(* IEC 61131-3 sources: Masterarbeit/sigmatek/lasalclass2/PW022_hardware/Class/SafetyManager (part 5) *)

END_FUNCTION

FUNCTION MyXSort VAR_INPUT p1:^void; p2:^void; END_VAR VAR_OUTPUT retcode : dint; END_VAR;

FUNCTION SafetyManager::MySort
  VAR_INPUT
    src 	: ^USINT;
    no 	: UDINT;
    itemsize 	: UDINT;
    sortfunct 	: ^void;
  END_VAR
  VAR_OUTPUT
    retcode 	: BOOL;
  END_VAR
  var
    tmp, hp : ^DINT;
    mx, nx, wx, parent, child, max, i : dint;
    spuf : array[0..127] of dint;
  end_var

  retcode := false;

  // work faster with the pointer list (no memcopy used)
  if itemsize = 4 then
    nx      := to_dint(no);
    mx      := (nx + 6) / 8;
    src     := src;
    tmp     := #spuf[0];
    retcode := true;

    while(1) do
      if(mx) then
        mx     -= 1;
        parent := mx;
        tmp^ := (src$^DINT + (parent$udint*4))^;
      else
        nx -= 1;
        if(nx) then
          hp := src + (nx$udint*4);
          tmp^ := hp^;
          hp^ := (src$^DINT)^;
          parent := 0;
        else
          exit;
        end_if;
      end_if;

      child := parent * 8 + 1;
      while(child < nx) do
        wx := nx - child;
        if(wx > 8) then
          wx := 8;
        end_if;

        max := 0;
        if(wx > 1) then
          for i:=1 to wx-1 do
            if(sortfunct$MyXSort(src+(to_udint(child+i)*4), src+to_udint(child+max)*4) > 0) then
              max := i;
            end_if;
          end_for;
        end_if;

        child += max;

        if(sortfunct$MyXSort(src+(child$udint*4), tmp) <= 0) then
          exit;
        end_if;

        (src$^DINT+(parent$udint*4))^ := (src$^DINT+(child$udint*4))^;
        parent := child;
        child  := parent * 8 + 1;
      end_while;

      (src$^DINT+(parent$udint*4))^ := tmp^;
    end_while;
  else
    if(itemsize <= sizeof(spuf)) then

      nx      := to_dint(no);
      mx      := (nx + 6) / 8;
      src     := src;
      tmp     := #spuf[0];
      retcode := true;

      while(1) do
        if(mx) then
          mx     -= 1;
          parent := mx;
          _memcpy(tmp, src + (parent$udint*itemsize), itemsize);
        else
          nx -= 1;
          if(nx) then
            hp := src + (nx$udint*itemsize);
            _memcpy(tmp, hp, itemsize);
            _memmove(hp, src, itemsize);
            parent := 0;
          else
            exit;
          end_if;
        end_if;

        child := parent * 8 + 1;
        while(child < nx) do
          wx := nx - child;
          if(wx > 8) then
            wx := 8;
          end_if;

          max := 0;
          if(wx > 1) then
            for i:=1 to wx-1 do
              if(sortfunct$MyXSort(src+(to_udint(child+i)*itemsize), src+to_udint(child+max)*itemsize) > 0) then
                max := i;
              end_if;
            end_for;
          end_if;

          child += max;

          if(sortfunct$MyXSort(src+(child$udint*itemsize), tmp) <= 0) then
            exit;
          end_if;

          _memcpy(src+(parent$udint*itemsize), src+(child$udint*itemsize), itemsize);
          parent := child;
          child  := parent * 8 + 1;
        end_while;

        _memcpy(src+(parent$udint*itemsize), tmp, itemsize);
      end_while;
    end_if;
  end_if;

END_FUNCTION

FUNCTION SafetyManager::ConnectionSort
  VAR_INPUT
    pCon1 	: ^pVoid;
    pCon2 	: ^pVoid;
  END_VAR
  VAR_OUTPUT
    retcode 	: DINT;
  END_VAR
  VAR
    Var1 : HDINT;
    Var2 : HDINT;
    pHelp : ^HDINT;
    Uint1 : UINT;
    Uint2 : UINT;
  END_VAR

  // dint MyXSort(void *p1, void *p2)
  //   if(a>b) retcode = 1;
  //   if(a=b) retcode = 0;
  //   if(a<b) retcode = -1

  pHelp := (pCon1^$^t_FSoEConnectionDetails^.pSlavePathComp)$^HDINT;
  if pHelp then
    if pHelp^$USINT = INTERFACE_CRC_MODE then
      Var1 := (pHelp + 1)^;
    else
      // no interface frame => sort to the end
      Var1 := 16#FFFFFFFF;
    end_if;
  else
    // no compressed path available => sort to the end
    Var1 := 16#FFFFFFFF;
  end_if;

  pHelp := (pCon2^$^t_FSoEConnectionDetails^.pSlavePathComp)$^HDINT;
  if pHelp then
    if pHelp^$USINT = INTERFACE_CRC_MODE then
      Var2 := (pHelp + 1)^;
    else
      // no interface frame => sort to the end
      Var2 := 16#FFFFFFFF;
    end_if;
  else
    // no compressed path available => sort to the end
    Var2 := 16#FFFFFFFF;
  end_if;

  // we want all connections to be sorted by the Interface CRC
  if Var1 > Var2 then
    retcode := 1;
  elsif Var1 < Var2 then
    retcode := -1;
  else
    // not possible with unique Interface CRCs, but a slave can provide between 1 and 150 connections with the same settings (only different offsets)
    // therefore it can only be detected as an error if the sources differ and they are not interface masters
    if pCon1^$^t_FSoEConnectionDetails^.OwnerSafetyNbr <> pCon2^$^t_FSoEConnectionDetails^.OwnerSafetyNbr then
      retcode := 0;
    else
      // otherwise sort by offset
      Uint1 := pCon1^$^t_FSoEConnectionDetails^.SlaveReadOffset;
      Uint2 := pCon2^$^t_FSoEConnectionDetails^.SlaveReadOffset;

      if Uint1 > Uint2 then
        retcode := 1;
      elsif Uint1 < Uint2 then
        retcode := -1;
      else
        retcode := 0;
      end_if;
    end_if;
  end_if;

END_FUNCTION

FUNCTION SafetyManager::FinalizePDOMapping
  VAR
    pHelpConnection   : ^t_FSoEConnectionDetails;
    pHelpSafety       : ^t_SafetyComponent;
    i                 : UDINT;
    ModuleReadOffset  : UINT;
    ModuleReadSize    : UINT;
    ModuleWriteOffset : UINT;
    ModuleWriteSize   : UINT;
    MngReadOffset     : UINT;
    MngReadSize       : UINT;
    MngWriteOffset    : UINT;
    MngWriteSize      : UINT;
    MyPara            : CmdStruct;
    MyResult          : results;
    bIsCustomConnValid: BOOL;
  END_VAR

  // check the FSoE Infos from the other side
  if IFFSoENo then
    for i := 0 to (IFFSoENo-1) do
      // search for a local module to handle this
      pHelpConnection := pSortedConnections;
      while pHelpConnection do
        bIsCustomConnValid := CheckCustomConnectionValid(pHelpConnection,#aIFFSoEInfos[i]);
        if (bIsCustomConnValid                    |
           ((pHelpConnection^.SlaveAddress)  &
           (pHelpConnection^.SlaveAddress    =  aIFFSoEInfos[i].FromOtherSide.SlaveAddress)))  &
           (pHelpConnection^.Flags.IsMaster  <> aIFFSoEInfos[i].FromOtherSide.Flags.IsMaster)  &
           (pHelpConnection^.MasterReadSize  =  aIFFSoEInfos[i].FromOtherSide.MasterReadSize)  &
           (pHelpConnection^.MasterWriteSize =  aIFFSoEInfos[i].FromOtherSide.MasterWriteSize) &
           (pHelpConnection^.InternalConnectionState =  FCS_RESET) then

          // now we check the interface CRC
          if pHelpConnection^.pSlavePathComp & pHelpConnection^.SlavePathCompLen then
            if aIFFSoEInfos[i].FromOtherSide.InterfaceCRC = (pHelpConnection^.pSlavePathComp$^HDINT + 1)^ then
              pHelpSafety := pFirstSafetyComponent;
              while pHelpSafety do
                if pHelpSafety^.SafetyNbr = pHelpConnection^.OwnerSafetyNbr then
                  exit;
                end_if;

                pHelpSafety := pHelpSafety^.pNext;
              end_while;

              if pHelpSafety then
                if pHelpConnection^.Flags.IsMaster then
#ifdef SAFETY_DEBUG_LOGGING_ACTIVATED
#pragma message("RamAnd 20.11.2014 16:41 \ testweise mapping loggen")
                  LogValue("@DBG (SafetyManager::FinalizePDOMapping) <This side is Master> ConnectionID: 0x{0}, SlaveAddress: 0x{1}, InterfaceCRC: 0x{2}", Value:=pHelpConnection^.ConnectionID, Value2:=pHelpConnection^.SlaveAddress, Value3 := aIFFSoEInfos[i].FromOtherSide.InterfaceCRC);
#endif

                  // the module is master and the managing module slave
                  ModuleReadOffset  := pHelpConnection^.MasterReadOffset;
                  ModuleReadSize    := pHelpConnection^.MasterReadSize;
                  ModuleWriteOffset := pHelpConnection^.MasterWriteOffset;
                  ModuleWriteSize   := pHelpConnection^.MasterWriteSize;
                  MngReadOffset     := 0; // offsets in managing modules are always dynamic
                  MngReadSize       := pHelpConnection^.MasterWriteSize;
                  MngWriteOffset    := 0; // offsets in managing modules are always dynamic
                  MngWriteSize      := pHelpConnection^.MasterReadSize;
                else
#ifdef SAFETY_DEBUG_LOGGING_ACTIVATED
#pragma message("RamAnd 20.11.2014 16:41 \ testweise mapping loggen")
                  LogValue("@DBG (SafetyManager::FinalizePDOMapping) <This side is Slave> ConnectionID: 0x{0}, SlaveAddress: 0x{1}, InterfaceCRC: 0x{2}", Value:=aIFFSoEInfos[i].FromOtherSide.ConnectionID, Value2:=aIFFSoEInfos[i].FromOtherSide.SlaveAddress, Value3 := aIFFSoEInfos[i].FromOtherSide.InterfaceCRC);
#endif

                  // the module is slave and the managing module master
                  ModuleReadOffset  := pHelpConnection^.SlaveReadOffset;
                  ModuleReadSize    := pHelpConnection^.MasterWriteSize;
                  ModuleWriteOffset := pHelpConnection^.SlaveWriteOffset;
                  ModuleWriteSize   := pHelpConnection^.MasterReadSize;
                  MngReadOffset     := 0; // offsets in managing modules are always dynamic
                  MngReadSize       := pHelpConnection^.MasterReadSize;
                  MngWriteOffset    := 0; // offsets in managing modules are always dynamic
                  MngWriteSize      := pHelpConnection^.MasterWriteSize;
                end_if;

                MyPara.uiCmd := CMD_SM_ADD_OUTPUT_PDO;
                MyPara.aPara[0] := 1;  // mark as interface frame PDO
                pHelpSafety^.pThis^.NewInst(#MyPara, #MyResult);

//                  pPDOElement^.SourceInfo.pPDOMem       := MyResult.aData[0]$^USINT;
//                  pPDOElement^.SourceInfo.pPDOMemDPRAM  := MyResult.aData[4]$^USINT;
//                  pPDOElement^.SourceInfo.HandlePDODPRAM:= MyResult.aData[8]$UDINT;   // Needed for Payload Support
//                  pPDOElement^.SourceInfo.OffsetPDODPRAM:= MyResult.aData[12]$UDINT;  // Needed for Payload Support

                if FSoECopyCmdNo < MAX_FSOE_CONNECTIONS then
                  aFSoECopyCmds[FSoECopyCmdNo].pSource  := MyResult.aData[0]$^USINT + ModuleReadOffset;
                  aFSoECopyCmds[FSoECopyCmdNo].pDest    := aIFFSoEInfos[i].pManaging^.pPDOWriteSpace + aIFFSoEInfos[i].pManaging^.PDOWriteMemUsed;
                  aFSoECopyCmds[FSoECopyCmdNo].Size     := ModuleReadSize;
                  FSoECopyCmdNo                         += 1;
                else
                  LogValue("@0493 (SafetyManager::FinalizePDOMapping) Maximum limit of allowed FSoE connections exceeded (0x{0})", Value:=MAX_FSOE_CONNECTIONS);
                end_if;

#ifdef SAFETY_DEBUG_LOGGING_ACTIVATED
#pragma message("RamAnd 20.11.2014 16:41 \ testweise mapping loggen")
                LogValue("@DBG (SafetyManager::FinalizePDOMapping) Modul => Mng: Rd Offset Modul: 0x{0}, Wr Offset Mng: 0x{1}, Größe: 0x{2}", Value:=ModuleReadOffset, Value2:=aIFFSoEInfos[i].pManaging^.PDOWriteMemUsed, Value3:=ModuleReadSize);
#endif

                aIFFSoEInfos[i].pManaging^.PDOWriteMemUsed += MngWriteSize;

                MyPara.uiCmd := CMD_SM_PDO_MEM_USAGE_WR;
                MyPara.aPara[0] := aIFFSoEInfos[i].pManaging^.PDOWriteMemUsed$DINT;
                aIFFSoEInfos[i].pManaging^.pThis^.NewInst(#MyPara, #MyResult);

                MyPara.uiCmd := CMD_SM_ADD_INPUT_PDO;
                MyPara.aPara[0] := (aIFFSoEInfos[i].pManaging^.pPDOReadSpace + aIFFSoEInfos[i].pManaging^.PDOReadMemUsed)$DINT;
                MyPara.aPara[1] := 0;
                MyPara.aPara[2] := aIFFSoEInfos[i].FromOtherSide.SafetyNbr$DINT;
                MyPara.aPara[3] := ModuleWriteSize;
                MyPara.aPara[4] := 0;
                MyPara.aPara[5] := 0;
                MyPara.aPara[6] := 0;
                MyPara.aPara[7] := ModuleWriteOffset;
                MyPara.aPara[8] := SM_IF_VALIDITY_MARK$DINT;
                MyPara.aPara[9] := TRUE;

                pHelpSafety^.pThis^.NewInst(#MyPara, #MyResult);

                if FSoEInputPDONo < MAX_FSOE_CONNECTIONS then
                  aFSoEInputPDOs[FSoEInputPDONo].pSafety    := pHelpSafety;
                  aFSoEInputPDOs[FSoEInputPDONo].pMem       := MyPara.aPara[0];
                  FSoEInputPDONo += 1;
                else
                  LogValue("@0490 (SafetyManager::FinalizePDOMapping) Maximum limit of allowed FSoE input Frames exceeded (0x{0})", Value:=MAX_FSOE_CONNECTIONS);
                end_if;

#ifdef SAFETY_DEBUG_LOGGING_ACTIVATED
#pragma message("RamAnd 20.11.2014 16:41 \ testweise mapping loggen")
                LogValue("@DBG (SafetyManager::FinalizePDOMapping) Mng => Modul: Wr Offset Modul: 0x{0}, Rd Offset Mng: 0x{1}, Größe: 0x{2}", Value:=ModuleWriteOffset, Value2:=aIFFSoEInfos[i].pManaging^.PDOReadMemUsed, Value3:=ModuleWriteSize);
#endif

                aIFFSoEInfos[i].pManaging^.PDOReadMemUsed += MngReadSize;

                MyPara.uiCmd := CMD_SM_PDO_MEM_USAGE_RD;
                MyPara.aPara[0] := aIFFSoEInfos[i].pManaging^.PDOReadMemUsed$DINT;
                aIFFSoEInfos[i].pManaging^.pThis^.NewInst(#MyPara, #MyResult);

                // mark the connection as established
                pHelpConnection^.InternalConnectionState := FCS_CONNECTION;

                // we found something for this connection => continue with the next
                exit;
              else
                LogValue("@0495 (SafetyManager::FinalizePDOMapping) Could not find safety module with safety number 0x{0} for FSoE interface connection", Value:=pHelpConnection^.OwnerSafetyNbr);
              end_if;
            end_if;
          end_if;
        end_if;

        pHelpConnection := pHelpConnection^.pNextSorted;
      end_while;
    end_for;
  end_if;

END_FUNCTION

FUNCTION SafetyManager::AddInternalIFFSoE
  VAR_INPUT
    pMasterConnection 	: ^t_FSoEConnectionDetails;
    pMasterConfig 	: ^t_CfgListElem;
    pSlaveConnection 	: ^t_FSoEConnectionDetails;
    pSlaveConfig 	: ^t_CfgListElem;
  END_VAR
  VAR
    i             : USINT;
    InterfaceCRC  : HDINT;
    pHelpSafety   : ^t_SafetyComponent;
    pMasterSafety : ^t_SafetyComponent;
    pSlaveSafety  : ^t_SafetyComponent;
    MyPara 	      : CmdStruct;
    MyResult	    : results;
    pPDOReadData  : pVoid;
    AddToList     : BOOL;
  END_VAR

  if pMasterConnection^.pSlavePathComp then
    InterfaceCRC := (pMasterConnection^.pSlavePathComp$^HDINT + 1)^;
  else
    // no interface CRC available
    return;
  end_if;

  AddToList := TRUE;
  if LocalIFNo then
    // check if the interfaceCRCs are already registered
    for i := 0 to (LocalIFNo-1) do
      if (aLocalIFs[i].InterfaceCRC = InterfaceCRC) & (aLocalIFs[i].MasterSafetyNbr = pMasterConfig^.SafetyNbr) then
        // already in the list => leave to prevent adding a second time
        AddToList := FALSE;
        return;
      end_if;
    end_for;
  end_if;

  pSlaveSafety := NIL;

  pHelpSafety := pFirstSafetyComponent;
  while pHelpSafety do

    if pHelpSafety^.SafetyNbr = pSlaveConfig^.SafetyNbr then
      pSlaveSafety := pHelpSafety;
      exit;
    end_if;

    pHelpSafety := pHelpSafety^.pNext;
  end_while;

  if pSlaveSafety & AddToList then
    if LocalIFNo < MAX_INTERNAL_IF_MODULES then
      aLocalIFs[LocalIFNo].InterfaceCRC     := InterfaceCRC;
      aLocalIFs[LocalIFNo].pSafetyModule    := pSlaveSafety;
       aLocalIFs[LocalIFNo].MasterSafetyNbr := pMasterConfig^.SafetyNbr;
      LocalIFNo                           += 1;
    else
      LogValue("@0496 (SafetyManager::ShareConnectionInfos) Maximum limit of allowed local FSoE connections exceeded (0x{0})", Value:=MAX_INTERNAL_IF_MODULES);
    end_if;
  end_if;

//*****************************************************************************
//** TELL THE MODULES WHAT DATA TO COPY IN REALTIME                          **
//*****************************************************************************

  pMasterSafety  := NIL;

  pHelpSafety := pFirstSafetyComponent;
  while pHelpSafety do

    if pHelpSafety^.SafetyNbr = pMasterConfig^.SafetyNbr then
      pMasterSafety := pHelpSafety;
      exit;
    end_if;

    pHelpSafety := pHelpSafety^.pNext;
  end_while;

  // if we found the safety modules who are keeping the configs => tell them what to copy
  if pMasterSafety & pSlaveSafety then
    // check for equal sizes
    if (pMasterConnection^.MasterReadSize <> pSlaveConnection^.MasterReadSize) |
       (pMasterConnection^.MasterWriteSize <> pSlaveConnection^.MasterWriteSize) then
      LogValue("@048E (SafetyManager::ShareConnectionInfos) Error! The sizes of master and slave connection do not match for Slave Address 0x{0} and ConnectionID 0x{1}!", Value:=pMasterConnection^.SlaveAddress, Value2:=pMasterConnection^.ConnectionID);
      return;
    end_if;

    // we start with the safe outputs: get the data pointer from the master and give it to the slave
    MyPara.uiCmd    := CMD_SM_ADD_OUTPUT_PDO;
    MyResult.uiLng  := 0;
    pMasterSafety^.pThis^.NewInst(#MyPara, #MyResult);

    if MyResult.uiLng <> 4 then
      LogError("@048F (SafetyManager::ShareConnectionInfos) Invalid return value when asking the master safety module for it's pointer to the PDO read data!");
      return;
    end_if;

    pPDOReadData := MyResult.aData[0]$pVoid;

#ifdef SAFETY_DEBUG_LOGGING_ACTIVATED
#pragma message("RamAnd 20.11.2014 16:41 \ testweise mapping loggen")
    LogValue("@DBG (SafetyManager::AddInternalIFFSoE) ConnectionID: {0}, SlaveAddress: {1}, InterfaceCRC: {2}", Value:=pMasterConnection^.ConnectionID, Value2:=pMasterConnection^.SlaveAddress, Value3 := InterfaceCRC);
    LogValue("@DBG (SafetyManager::AddInternalIFFSoE) MasterSafetyNbr: {0}, SlaveSafetyNbr: {1}", Value:=pMasterConnection^.OwnerSafetyNbr, Value2:=pSlaveConnection^.OwnerSafetyNbr);
    LogValue("@DBG (SafetyManager::AddInternalIFFSoE) MasterReadOffset: {0}, MasterReadSize: {1}, SlaveWriteOffset: {2}", Value:=pMasterConnection^.MasterReadOffset, Value2:=pMasterConnection^.MasterReadSize, Value3 := pSlaveConnection^.SlaveWriteOffset);
#endif

    MyPara.uiCmd    := CMD_SM_ADD_INPUT_PDO;
    MyPara.aPara[0] := pPDOReadData$DINT + pMasterConnection^.MasterReadOffset;
    MyPara.aPara[2] := pMasterConnection^.OwnerSafetyNbr$DINT;
    MyPara.aPara[3] := pMasterConnection^.MasterReadSize;
    MyPara.aPara[4] := pMasterSafety^.InfoBits.IsOptional;
    MyPara.aPara[7] := pSlaveConnection^.SlaveWriteOffset;
    MyPara.aPara[8] := SM_IF_VALIDITY_MARK$DINT;
    MyPara.aPara[9] := TRUE;
    pSlaveSafety^.pThis^.NewInst(#MyPara, #MyResult);

    if FSoEInputPDONo < MAX_FSOE_CONNECTIONS then
      aFSoEInputPDOs[FSoEInputPDONo].pSafety    := pSlaveSafety;
      aFSoEInputPDOs[FSoEInputPDONo].pMem       := MyPara.aPara[0];
      FSoEInputPDONo += 1;
    else
      LogValue("@0490 (SafetyManager::AddInternalIFFSoE) Maximum limit of allowed FSoE input Frames exceeded (0x{0})", Value:=MAX_FSOE_CONNECTIONS);
    end_if;

    // safe inputs: get the data pointer from the slave and give it to the master
    MyPara.uiCmd    := CMD_SM_ADD_OUTPUT_PDO;
    MyResult.uiLng  := 0;
    pSlaveSafety^.pThis^.NewInst(#MyPara, #MyResult);

    if MyResult.uiLng <> 4 then
      LogError("@0491 (SafetyManager::AddInternalIFFSoE) Invalid return value when asking the slave safety module for it's pointer to the PDO read data!");
      return;
    end_if;

    pPDOReadData := MyResult.aData[0]$pVoid;

#ifdef SAFETY_DEBUG_LOGGING_ACTIVATED
#pragma message("RamAnd 20.11.2014 16:41 \ testweise mapping loggen")
    LogValue("@DBG (SafetyManager::AddInternalIFFSoE) SlaveReadOffset: {0}, SlaveReadSize: {1}, MasterWriteOffset: {2}", Value:=pSlaveConnection^.SlaveReadOffset, Value2:=pMasterConnection^.MasterWriteSize, Value3 := pMasterConnection^.MasterWriteOffset);
#endif

    MyPara.uiCmd    := CMD_SM_ADD_INPUT_PDO;
    MyPara.aPara[0] := pPDOReadData$DINT + pSlaveConnection^.SlaveReadOffset;
    MyPara.aPara[2] := pSlaveConnection^.OwnerSafetyNbr$DINT;
    MyPara.aPara[3] := pMasterConnection^.MasterWriteSize;
    MyPara.aPara[4] := pSlaveSafety^.InfoBits.IsOptional;
    MyPara.aPara[7] := pMasterConnection^.MasterWriteOffset;
    MyPara.aPara[8] := SM_IF_VALIDITY_MARK$DINT;
    MyPara.aPara[9] := TRUE;
    pMasterSafety^.pThis^.NewInst(#MyPara, #MyResult);

    if FSoEInputPDONo < MAX_FSOE_CONNECTIONS then
      aFSoEInputPDOs[FSoEInputPDONo].pSafety    := pMasterSafety;
      aFSoEInputPDOs[FSoEInputPDONo].pMem       := MyPara.aPara[0];
      FSoEInputPDONo += 1;
    else
      LogValue("@0490 (SafetyManager::AddInternalIFFSoE) Maximum limit of allowed FSoE input Frames exceeded (0x{0})", Value:=MAX_FSOE_CONNECTIONS);
    end_if;

    pSlaveConnection^.InternalConnectionState   := FCS_CONNECTION;

    // for easier debugging we take the values to the manager-connection as well (only for debugging to have the correct values in the connections)
    pMasterConnection^.InternalConnectionState  := FCS_CONNECTION;
    pMasterConnection^.SlaveReadOffset          := pSlaveConnection^.SlaveReadOffset;
    pMasterConnection^.SlaveWriteOffset         := pSlaveConnection^.SlaveWriteOffset;
  end_if;

END_FUNCTION

FUNCTION SafetyManager::CheckOptional
  VAR
    pHelpConfig     : ^t_CfgListElem;
    pHelpConfig2    : ^t_CfgListElem;
    pHelpSlaveCfg   : ^t_SlaveListElem;
    pHelpModuleCfg  : ^t_ModuleListElem;
    FoundIt         : BOOL;
  END_VAR

  // check all available configs
  pHelpConfig := pConfigs;
  while pHelpConfig do

    // search in module configs
    pHelpModuleCfg := pHelpConfig^.pFirstModuleCfg;
    while pHelpModuleCfg do
      if pHelpModuleCfg^.ModuleInfo.Info.IsOptional = FALSE then
        // if the slave config is not optional => check if we got the config
        FoundIt := FALSE;
        pHelpConfig2 := pConfigs;
        while pHelpConfig2 & (FoundIt = FALSE) do
          if (pHelpConfig2^.pFirstModuleCfg^.ModuleInfo.PathLen = pHelpModuleCfg^.ModuleInfo.PathLen) &
             (_memcmp(ptr1:=pHelpConfig2^.pFirstModuleCfg^.ModuleInfo.pPath, ptr2:=pHelpModuleCfg^.ModuleInfo.pPath, cntr:=pHelpModuleCfg^.ModuleInfo.PathLen) = 0) then

            FoundIt := TRUE;
            exit;
          end_if;

          pHelpConfig2 := pHelpConfig2^.pNext;
        end_while;

        if FoundIt = FALSE then
          // non-optional config not available
          return;
        end_if;
      end_if;

      pHelpModuleCfg := pHelpModuleCfg^.pNext;
    end_while;

    // search in slave configs
    pHelpSlaveCfg := pHelpConfig^.pFirstSlaveCfg;
    while pHelpSlaveCfg do
      if pHelpSlaveCfg^.SlaveInfo.Info.IsOptional = FALSE then
        // if the slave config is not optional => check if we got the config
        FoundIt := FALSE;
        pHelpConfig2 := pConfigs;
        while pHelpConfig2 do
          if pHelpConfig2^.pFirstModuleCfg & (pHelpConfig2^.pFirstModuleCfg^.ModuleInfo.PathLen = pHelpSlaveCfg^.SlaveInfo.PathLen) &
             (_memcmp(ptr1:=pHelpConfig2^.pFirstModuleCfg^.ModuleInfo.pPath, ptr2:=pHelpSlaveCfg^.SlaveInfo.pPath, cntr:=pHelpSlaveCfg^.SlaveInfo.PathLen) = 0) then

            FoundIt := TRUE;
            exit;
          end_if;

          pHelpConfig2 := pHelpConfig2^.pNext;
        end_while;

        if FoundIt = FALSE then
          // non-optional config not available
          return;
        end_if;
      end_if;

      pHelpSlaveCfg := pHelpSlaveCfg^.pNext;
    end_while;

    pHelpConfig := pHelpConfig^.pNext;
  end_while;

  // if nothing non-optional is missing => we're good to go (if something would be missing the method would have been left at this position)
  b_MandatoryStuffAvailable := TRUE;

END_FUNCTION

FUNCTION SafetyManager::FSoEConInitialized
  VAR_INPUT
    SafetyNbr 	: HDINT;
    ConnectionNo 	: UDINT;
    pFirstConnection 	: ^t_FSoEConnectionDetails;
  END_VAR
  VAR
    i               : UDINT;
    pActConnection  : ^t_FSoEConnectionDetails;
    pActConnLocal   : ^t_FSoEConnectionDetails;
    pHelpConfig     : ^t_CfgListElem;
  END_VAR

  // search for the configuration of the safety component
  pHelpConfig := pConfigs;
  while pHelpConfig do
    if pHelpConfig^.SafetyNbr = SafetyNbr then
      // found the module => now update the connection infos
      pActConnLocal  := pHelpConfig^.pFirstFSoEConnection;
      pActConnection := pFirstConnection;
      for i := 0 to (ConnectionNo-1) do
        // no valid local connection => leave
        if pActConnLocal = NIL then
          return;
        end_if;

        if pActConnLocal^.ConnectionState = FCS_NOT_INITIALIZED then
          // update slave address first because we are in background here and the data is also accessed in cyclic (connection state is checked first in cyclic)
          pActConnLocal^.SlaveAddress := pActConnection^.SlaveAddress;

          // now update the connection state
          pActConnLocal^.ConnectionState := pActConnection^.ConnectionState;
        end_if;

        pActConnLocal  := pActConnLocal^.pNext;
        pActConnection += sizeof(t_FSoEConnectionDetails);
      end_for;
    end_if;

    pHelpConfig := pHelpConfig^.pNext;
  end_while;

  CheckLocalSlaveAddresses();

  if InitSSW = _InitFinished then
    // maybe we have some new informations here
    CreateFSoEPDOs();
  end_if;

END_FUNCTION

FUNCTION SafetyManager::CheckLocalSlaveAddresses
  VAR
    pActConnection  : ^t_FSoEConnectionDetails;
    pHelpConfig     : ^t_CfgListElem;
  END_VAR

  // check if we got all slave addresses
  pHelpConfig := pConfigs;
  while pHelpConfig do
    pActConnection := pHelpConfig^.pFirstFSoEConnection;
    while pActConnection do
      if (pActConnection^.ConnectionState = FCS_NOT_INITIALIZED) then
        // as soon as we find a not initialized connection => leave
        return;
      end_if;

      pActConnection := pActConnection^.pNext;
    end_while;

    pHelpConfig := pHelpConfig^.pNext;
  end_while;

  // if we got this far, we got all slave addresses
  b_AllLocalSlaveAddressesValid := TRUE;

END_FUNCTION

FUNCTION SafetyManager::AddUdpConnection
  VAR_INPUT
    IP 	: HDINT;
    IFCRC 	: HDINT;
    SafetyNumber 	: HDINT;
    ProducerList 	: BOOL;
    ppConnection 	: ^t_pUdpConnection;(* := NIL *)
  END_VAR
  VAR_OUTPUT
    success 	: BOOL;
  END_VAR
  VAR
    i : UDINT;
    pActConnection : ^t_UdpConnection;
  END_VAR

  success := FALSE;

  // if we're consumer we add the connection to the producer list, because it's our producer
  if ProducerList then
    if sUdpVars.paConnectionsToProducers = NIL then
      bd_LogRtMessagesInCy.UdpNoMem4Connections := TRUE;
      return;
    end_if;

    // check if it already exists
    if sUdpVars.ProducerConnectionNo then
      pActConnection := #sUdpVars.paConnectionsToProducers^[0];
      for i := 0 to (sUdpVars.ProducerConnectionNo-1) do
        // we only add a new connection if it doesn't exist yet
        if (pActConnection^.IP = IP) & (pActConnection^.IFCRC = IFCRC) then
          // already existing
          LogValue("@0499 (SafetyManager::AddUdpConnection) Found 2 equal producer connections (IP: 0x{0}, IF CRC: 0x{1}) which is not possible to handle", Value:=IP, Value2:=IFCRC);
          return;
        end_if;
        pActConnection += sizeof(t_UdpConnection);
      end_for;
    end_if;

    pActConnection := #sUdpVars.paConnectionsToProducers^[sUdpVars.ProducerConnectionNo];

    pActConnection^.IP                            := IP;
    pActConnection^.IFCRC                         := IFCRC;
    pActConnection^.SafetyNbr                     := SafetyNumber;

    // reset some elements
    pActConnection^.SafetyNbrOtherSide            := 0;
    pActConnection^.InfoBits                      := 0;
    pActConnection^.WaitForResponse               := FALSE;
    pActConnection^.SendResponse                  := FALSE;
    pActConnection^.bSequenceCntReceived          := FALSE; //reset flag to allow sequence counter for new udp communication
    pActConnection^.ActReceiveData.usHeaderVersion := 0;
    pActConnection^.ActSendData.usHeaderVersion    := 0;
    pActConnection^.SentPackages                   := 0;
    pActConnection^.ReceivedPackages               := 0;
    pActConnection^.MaxResponseTime                := 0;
    pActConnection^.ActSendData.PdoLength          := 0;
    pActConnection^.ActSendData.SdoLength          := 0;
    pActConnection^.ActReceiveData.PdoLength       := 0;
    pActConnection^.ActReceiveData.SdoLength       := 0;
    sUdpVars.ProducerConnectionNo                   += 1;
    success                                         := TRUE;

    if ppConnection then
      ppConnection^ := pActConnection;
    end_if;
  else
    if sUdpVars.paConnectionsToConsumers = NIL then
      bd_LogRtMessagesInCy.UdpNoMem4Connections   := TRUE;
      return;
    end_if;

    // check if it already exists
    if sUdpVars.ConsumerConnectionNo then
      pActConnection := #sUdpVars.paConnectionsToConsumers^[0];
      for i := 0 to (sUdpVars.ConsumerConnectionNo-1) do
        // we only add a new connection if it doesn't exist yet
        if (pActConnection^.IP = IP) & (pActConnection^.IFCRC = IFCRC) then
          // already existing
          LogValue("@049A (SafetyManager::AddUdpConnection) Found 2 equal consumer connections (IP: 0x{0}, IF CRC: 0x{1}) which is not possible to handle", Value:=IP, Value2:=IFCRC);
          return;
        end_if;
        pActConnection += sizeof(t_UdpConnection);
      end_for;
    end_if;

    pActConnection := #sUdpVars.paConnectionsToConsumers^[sUdpVars.ConsumerConnectionNo];

    pActConnection^.IP                            := IP;
    pActConnection^.IFCRC                         := IFCRC;
    pActConnection^.SafetyNbr                     := SafetyNumber;

    // reset some elements
    pActConnection^.SafetyNbrOtherSide              := 0;
    pActConnection^.InfoBits                        := 0;
    pActConnection^.WaitForResponse                 := FALSE;
    pActConnection^.SendResponse                    := FALSE;
    pActConnection^.bSequenceCntReceived            := FALSE; //reset flag to allow sequence counter for new udp communication
    pActConnection^.ActReceiveData.usHeaderVersion  := 0;
    pActConnection^.ActSendData.usHeaderVersion     := 0;
    pActConnection^.SentPackages                    := 0;
    pActConnection^.ReceivedPackages                := 0;
    pActConnection^.MaxResponseTime                 := 0;
    pActConnection^.ActSendData.PdoLength           := 0;
    pActConnection^.ActSendData.SdoLength           := 0;
    pActConnection^.ActReceiveData.PdoLength        := 0;
    pActConnection^.ActReceiveData.SdoLength        := 0;

    sUdpVars.ConsumerConnectionNo                   += 1;
    success                                         := TRUE;

    if ppConnection then
      ppConnection^ := pActConnection;
    end_if;
  end_if;

  // whenever new connections are added, they need to be initialized
  sUdpVars.ConnectionsInitialized := FALSE;

END_FUNCTION

FUNCTION SafetyManager::UdpRequestScheduler
  VAR
    pActRequestEntry  : ^t_UdpConnection;
    pActRetryEntry    : ^t_UdpConnection;
    tmpretcode        : DINT;
    i                 : UDINT;
  END_VAR

  //point to actual request-entry
  pActRequestEntry := #sUdpVars.paConnectionsToProducers^[sUdpVars.RequestScheduler.ActRequestedIndex];

  //send a request every
  if ((sUdpVars.RequestScheduler.CyCnt MOD sUdpVars.CalculatedRequestTime) = 0) then
    //calculate actual time diff from last request to this
    sUdpVars.ActTimeRequestScheduler := ops.tAbsolute - sUdpVars.LastRequestTimeScheduler;
    sUdpVars.LastRequestTimeScheduler := ops.tAbsolute;

    //set maximal time diff of request scheduler call.
    if sUdpVars.MaxTimeRequestScheduler < sUdpVars.ActTimeRequestScheduler then
      sUdpVars.MaxTimeRequestScheduler := sUdpVars.ActTimeRequestScheduler;

      if sUdpVars.bSetFirstMaxRequestSchedulerTime = FALSE then
        //set initial value for time measure of maximum of request scheduler
        sUdpVars.bSetFirstMaxRequestSchedulerTime := TRUE;
        sUdpVars.MaxTimeRequestScheduler          := 0;
      end_if;
    end_if;

    // search through the list if something has to be sent (check also for changes in the data)
    for i := 0 to sUdpVars.ProducerConnectionNo-1 do

      //only send a request if not waiting for a response and the IP is valid (on cleaning out the connections some may be set to 0)
      if (pActRequestEntry^.WaitForResponse = FALSE) & (pActRequestEntry^.IP <> 0) then

        //send request to mover of actual entry
        tmpretcode := SendUdpRequest(pActRequestEntry);
        if tmpretcode >= 0 then

          //if sending was successful we are waiting for a response
          pActRequestEntry^.WaitForResponse   := TRUE;
          pActRequestEntry^.TLastRequest      := ops.tAbsolute;
          pActRequestEntry^.RequestRetries    := 0;

        else
          //unable to send request
          if bd_SingleLog.SendUdpReqFailed = FALSE then
            bd_SingleLog.SendUdpReqFailed := TRUE;
            LogError("@049B (SafetyManager::UdpRequestScheduler) [SL] Failed to send udp request");
          end_if;
        end_if;
      end_if;

      //increase actual index
      if sUdpVars.RequestScheduler.ActRequestedIndex < (sUdpVars.ProducerConnectionNo-1) then
        sUdpVars.RequestScheduler.ActRequestedIndex += 1;
      else
        // check the time of the cycle
        UdpSetTimeMeasurement();

        //when reaching last entry -> reset index
        sUdpVars.RequestScheduler.ActRequestedIndex := 0;
      end_if;

      pActRequestEntry := #sUdpVars.paConnectionsToProducers^[sUdpVars.RequestScheduler.ActRequestedIndex];
    end_for;

  // between the normal requests we do the retries
  elsif ((sUdpVars.RequestScheduler.CyCnt MOD UDP_RETRY_TIME) = 0) then

    pActRetryEntry := #sUdpVars.paConnectionsToProducers^[0];

    // check if we have to send a retry
    for i := 0 to sUdpVars.ProducerConnectionNo-1 do

      // look if we actual wait for a response to send retries and check if we didn't receive data in time
      if (pActRetryEntry^.WaitForResponse = TRUE) & ((ops.tAbsolute - pActRetryEntry^.TLastRequest) > sUdpVars.CalculatedRequestTimeout) then
        //check for connection timeout
        if (ops.tAbsolute-pActRetryEntry^.TLastValidRequest) > (UDP_DEFAULT_TRANSMISSION_TIME*2) then
          //reset header version if connection timeout is reached.
          pActRetryEntry^.ActReceiveData.usHeaderVersion := 0;
          pActRetryEntry^.ActSendData.usHeaderVersion    := 0;
          pActRetryEntry^.TLastValidRequest := ops.tAbsolute;
        end_if;

        if pActRetryEntry^.RequestRetries >= UDP_MAX_RETRIES then

          pActRetryEntry^.MaxRetryCnt     += 1;
          pActRetryEntry^.WaitForResponse := FALSE;

          //check for new header version with extended sequence number (4Byte)
          if pActRetryEntry^.ActSendData.usHeaderVersion >= UDP_HEADER_VERSION_V2 then
            // we did not get our response => increase the sequence number for the next attempt
            pActRetryEntry^.ActSendData.udSequenceNumber += 1;
          else
            // we did not get our response => increase the sequence number for the next attempt
            pActRetryEntry^.ActSendData.usSequenceNumber += 1;
            pActRetryEntry^.ActSendData.udSequenceNumber := pActRetryEntry^.ActSendData.usSequenceNumber;
          end_if;

        // only if the IP is valid
        elsif (pActRetryEntry^.IP <> 0) then

          //send retry to actual cpu
          tmpretcode := SendUdpRequest(pActRetryEntry);
          if tmpretcode >= 0 then
            pActRetryEntry^.TLastRequest   := ops.tAbsolute;
            pActRetryEntry^.RequestRetries += 1;
            exit;
          else
            //unable to send retry
            if bd_SingleLog.SendUdpReqRetryFailed = FALSE then
              bd_SingleLog.SendUdpReqRetryFailed := TRUE;
              LogError("@049D (SafetyManager::UdpTimeScheduler) [SL] Failed to send udp retry");
            end_if;
          end_if;
        end_if;

      end_if;

      pActRetryEntry += sizeof(t_UdpConnection);

    end_for;

  end_if;

  sUdpVars.RequestScheduler.CyCnt += 1;

END_FUNCTION

FUNCTION SafetyManager::UdpSetTimeMeasurement

  if sUdpVars.RequestScheduler.LastTime then
    sUdpVars.RequestScheduler.ActRuntime := ops.tAbsolute - sUdpVars.RequestScheduler.LastTime;
    if sUdpVars.RequestScheduler.ActRuntime > sUdpVars.RequestScheduler.MaxRuntime then
      sUdpVars.RequestScheduler.MaxRuntime := sUdpVars.RequestScheduler.ActRuntime;
    end_if;

    if sUdpVars.RequestScheduler.ActRuntime < sUdpVars.RequestScheduler.MinRuntime then
      sUdpVars.RequestScheduler.MinRuntime := sUdpVars.RequestScheduler.ActRuntime;
    end_if;
  else
    sUdpVars.RequestScheduler.MinRuntime := 9999;
  end_if;
  sUdpVars.RequestScheduler.LastTime := ops.tAbsolute;

END_FUNCTION

FUNCTION SafetyManager::SendUdpRequest
  VAR_INPUT
    pConnection 	: ^t_UdpConnection;
  END_VAR
  VAR_OUTPUT
    retcode 	: DINT;
  END_VAR
  VAR
    udActSendLength : UDINT;
  END_VAR

  sUdpVars.pTempSendBufferCy^.Header.Command   := t_UdpCommand::UdpCmd_DataReq;
  // add supported header version to state (is set if we got response from other side)
  sUdpVars.pTempSendBufferCy^.Header.State     := t_UdpPacketHeaderV2.State.IsFromConsumer + pConnection^.ActSendData.usHeaderVersion;
  sUdpVars.pTempSendBufferCy^.Header.IFCRC     := pConnection^.IFCRC;
  sUdpVars.pTempSendBufferCy^.Header.SafetyNbr := pConnection^.SafetyNbr;

  UdpSendData.SectionStart();

  //check for new header version with extended sequence number (4Byte)
  if pConnection^.ActSendData.usHeaderVersion >= UDP_HEADER_VERSION_V2 then

    sUdpVars.pTempSendBufferCy^.Header.SequenceNumber := pConnection^.ActSendData.udSequenceNumber;

    udActSendLength := sizeof(t_UdpPacketHeaderV2);

    if pConnection^.ActSendData.PdoLength then
      sUdpVars.pTempSendBufferCy^.Header.PdoDataLength  := pConnection^.ActSendData.PdoLength;
      _memcpy(ptr1:=#sUdpVars.pTempSendBufferCy^.Data, ptr2:=#pConnection^.ActSendData.PdoData, cntr:=pConnection^.ActSendData.PdoLength);
      udActSendLength += pConnection^.ActSendData.PdoLength;
    else
      sUdpVars.pTempSendBufferCy^.Header.PdoDataLength  := 0;
    end_if;

    if pConnection^.ActSendData.SdoLength then
      sUdpVars.pTempSendBufferCy^.Header.SdoDataLength  := pConnection^.ActSendData.SdoLength;
      _memcpy(ptr1:=#sUdpVars.pTempSendBufferCy^.Data + pConnection^.ActSendData.PdoLength, ptr2:=#pConnection^.ActSendData.SdoData, cntr:=pConnection^.ActSendData.SdoLength);
      udActSendLength += pConnection^.ActSendData.SdoLength;
    else
      sUdpVars.pTempSendBufferCy^.Header.SdoDataLength  := 0;
    end_if;

  else
    //use old headerversion with 1byte Sequence Counter
    sUdpVars.pTempSendBufferCy^$t_UdpPacketV1.Header.SequenceNumber := pConnection^.ActSendData.usSequenceNumber;

    udActSendLength := sizeof(t_UdpPacketHeaderV1);

    if pConnection^.ActSendData.PdoLength then
      sUdpVars.pTempSendBufferCy^$t_UdpPacketV1.Header.PdoDataLength  := pConnection^.ActSendData.PdoLength;
      _memcpy(ptr1:=#sUdpVars.pTempSendBufferCy^$t_UdpPacketV1.Data, ptr2:=#pConnection^.ActSendData.PdoData, cntr:=pConnection^.ActSendData.PdoLength);
      udActSendLength += pConnection^.ActSendData.PdoLength;
    else
      sUdpVars.pTempSendBufferCy^$t_UdpPacketV1.Header.PdoDataLength  := 0;
    end_if;

    if pConnection^.ActSendData.SdoLength then
      sUdpVars.pTempSendBufferCy^$t_UdpPacketV1.Header.SdoDataLength  := pConnection^.ActSendData.SdoLength;
      _memcpy(ptr1:=#sUdpVars.pTempSendBufferCy^$t_UdpPacketV1.Data + pConnection^.ActSendData.PdoLength, ptr2:=#pConnection^.ActSendData.SdoData, cntr:=pConnection^.ActSendData.SdoLength);
      udActSendLength += pConnection^.ActSendData.SdoLength;
    else
      sUdpVars.pTempSendBufferCy^$t_UdpPacketV1.Header.SdoDataLength  := 0;
    end_if;

  end_if;

  UdpSendData.SectionStop();

  retcode := SendUDPData(sUdpVars.pTempSendBufferCy, udActSendLength, pConnection^.IP);

  sUdpVars.SendCnt += 1;

  if retcode < 0 then
    // error at sending
    sUdpVars.LastSendError := retcode;
    sUdpVars.SendErrorCnt += 1;
  else
    // only send this once
    pConnection^.ActSendData.SdoLength := 0;

    pConnection^.SentPackages += 1;
  end_if;

END_FUNCTION

FUNCTION SafetyManager::ReceiveUdpData
  VAR_INPUT
    pData 	: ^void;
    udLength 	: UDINT;
    udIPAddr 	: HDINT;
    udPort 	: UDINT;
  END_VAR
  VAR
    i               : UDINT;
    FoundConnection : BOOL;
    pPacketHeader   : ^t_UdpPacketHeaderV2;
    pActConnection  : ^t_UdpConnection;
    pHelpCfg        : ^t_CfgListElem;
    pHelpModule     : ^t_ModuleListElem;
    retcode         : DINT;
  END_VAR

  pPacketHeader := pData$^t_UdpPacketHeaderV2;

  // only take the data if we're not clearing the routing infos at the very moment
  if InitSSW > _ClearRoutingInfos then

    // increase receive counter
    sUdpVars.ReceiveCnt += 1;

    // check for longest time between data packages
    if sUdpVars.LastReceivedTimeStamp then
      sUdpVars.ActTimeBetweenReceiveData := ops.tAbsolute - sUdpVars.LastReceivedTimeStamp;
      if sUdpVars.ActTimeBetweenReceiveData > sUdpVars.MaxTimeBetweenReceiveData then
        sUdpVars.MaxTimeBetweenReceiveData := sUdpVars.ActTimeBetweenReceiveData;
      end_if;
    end_if;
    sUdpVars.LastReceivedTimeStamp := ops.tAbsolute;

    if (pPacketHeader^.State AND (t_UdpFrameState.IsFromConsumer OR t_UdpFrameState.IsFromProducer)) = t_UdpFrameState.IsFromConsumer then
      // it's a request from a consumer => check our list of consumers

      // the only valid command here is data request
      if pPacketHeader^.Command = t_UdpCommand::UdpCmd_DataReq then
        FoundConnection := FALSE;
        if sUdpVars.ConsumerConnectionNo then
          pActConnection := #sUdpVars.paConnectionsToConsumers^[0];
          // check if it's one of our existing connections
          for i := 0 to sUdpVars.ConsumerConnectionNo-1 do
            if (pActConnection^.IP = udIPAddr) & (pActConnection^.SafetyNbrOtherSide = pPacketHeader^.SafetyNbr) then
              // check if it's the same IF CRC
              if (pActConnection^.IFCRC = pPacketHeader^.IFCRC) then
                FoundConnection := TRUE;
                exit;
              end_if;
            end_if;

            pActConnection += sizeof(t_UdpConnection);
          end_for;
        end_if;

        if FoundConnection then
          //check for new header version with extended sequence number (4Byte)
          if pData^$t_UdpPacketV2.Header.State and UDP_HEADER_VERSION_MASK >= UDP_HEADER_VERSION_V2 then
            // pActConnection points to the right connection
            HandleUdpRequestV2(pConnection:=pActConnection, pPacket:=pData$^t_UdpPacketV2, udLength:=udLength);
          else
            // pActConnection points to the right connection
            HandleUdpRequest(pConnection:=pActConnection, pPacket:=pData$^t_UdpPacketV1, udLength:=udLength);
          end_if;
          //set received header version
          pActConnection^.ActReceiveData.usHeaderVersion := (pData^$t_UdpPacketV2.Header.State and UDP_HEADER_VERSION_MASK);
          //we can set the headerversion from receive data also for the send data
          pActConnection^.ActSendData.usHeaderVersion    := pActConnection^.ActReceiveData.usHeaderVersion;
          //if we got header version info with version higher our own supported header version set the own supported version
          if pActConnection^.ActSendData.usHeaderVersion > UDP_HEADER_ACTVERSION then
            pActConnection^.ActSendData.usHeaderVersion := UDP_HEADER_ACTVERSION;
          end_if;
        else
          // search for the safety number of the producer
          pHelpCfg := pConfigs;
          while pHelpCfg do
            pHelpModule := pHelpCfg^.pFirstModuleCfg;
            while pHelpModule do
              if pHelpModule^.ModuleInfo.InterfaceCRC = pPacketHeader^.IFCRC then
                // add the connection (we're producer and we the consumer wants something from us)
                if AddUdpConnection(IP:=udIPAddr, IFCRC:=pPacketHeader^.IFCRC, SafetyNumber:=pHelpCfg^.SafetyNbr, ProducerList:=FALSE, #pActConnection) then
                  //check for new header version with extended sequence number (4Byte)
                  if pData^$t_UdpPacketV2.Header.State and UDP_HEADER_VERSION_MASK >= UDP_HEADER_VERSION_V2 then
                    // pActConnection points to the right connection
                    HandleUdpRequestV2(pConnection:=pActConnection, pPacket:=pData$^t_UdpPacketV2, udLength:=udLength);
                  else
                    // pActConnection points to the right connection
                    HandleUdpRequest(pConnection:=pActConnection, pPacket:=pData$^t_UdpPacketV1, udLength:=udLength);
                  end_if;
                  //set received header version
                  pActConnection^.ActReceiveData.usHeaderVersion := (pData^$t_UdpPacketV2.Header.State and UDP_HEADER_VERSION_MASK);
                  //we can set the headerversion from receive data also for the send data
                  pActConnection^.ActSendData.usHeaderVersion    := pActConnection^.ActReceiveData.usHeaderVersion;
                  //if we got header version info with version higher our own supported header version set the own supported version
                  if pActConnection^.ActSendData.usHeaderVersion > UDP_HEADER_ACTVERSION then
                    pActConnection^.ActSendData.usHeaderVersion := UDP_HEADER_ACTVERSION;
                  end_if;
                end_if;
                return;
              end_if;

              pHelpModule := pHelpModule^.pNext;
            end_while;

            pHelpCfg := pHelpCfg^.pNext;
          end_while;
          sUdpVars.UnhandledReceivePacketCnt += 1;
        end_if;

      else
        // invalid command
        bd_LogRtMessagesInCy.UdpReceivedInvalidCommand := TRUE;
        sUdpVars.UnhandledReceivePacketCnt += 1;
      end_if;
    elsif (pPacketHeader^.State AND (t_UdpFrameState.IsFromConsumer OR t_UdpFrameState.IsFromProducer)) = t_UdpFrameState.IsFromProducer then
      // it's a response from a producer => check our list of producers

      // the only valid command here is data response
      if pPacketHeader^.Command = t_UdpCommand::UdpCmd_DataRsp then

        if sUdpVars.ProducerConnectionNo then
          FoundConnection := FALSE;
          pActConnection := #sUdpVars.paConnectionsToProducers^[0];
          // check if it's one of our existing connections
          for i := 0 to sUdpVars.ProducerConnectionNo-1 do
            if (pActConnection^.IP = udIPAddr) & (pActConnection^.IFCRC = pPacketHeader^.IFCRC) then
              FoundConnection := TRUE;
              exit;
            end_if;

            pActConnection += sizeof(t_UdpConnection);
          end_for;

          if FoundConnection then
            //check for new version of udp header
            if pData^$t_UdpPacketV2.Header.State and UDP_HEADER_VERSION_MASK >= UDP_HEADER_VERSION_V2 then
              // pActConnection points to the right connection
              HandleUdpResponseV2(pConnection:=pActConnection, pPacket:=pData$^t_UdpPacketV2, udLength:=udLength);
            else
              // pActConnection points to the right connection
              HandleUdpResponse(pConnection:=pActConnection, pPacket:=pData$^t_UdpPacketV1, udLength:=udLength);
            end_if;
            pActConnection^.ActReceiveData.usHeaderVersion := pData^$t_UdpPacketV2.Header.State and UDP_HEADER_VERSION_MASK;
            //we can set the headerversion from receive data also for the send data
            pActConnection^.ActSendData.usHeaderVersion    := pActConnection^.ActReceiveData.usHeaderVersion;
            //if we got header version info with version higher our own supported header version set the own supported version
            if pActConnection^.ActSendData.usHeaderVersion > UDP_HEADER_ACTVERSION then
              pActConnection^.ActSendData.usHeaderVersion := UDP_HEADER_ACTVERSION;
            end_if;
          else
            // ignore it, maybe the safety project changed
            sUdpVars.UnhandledReceivePacketCnt += 1;
          end_if;

        else
          // ignore it, maybe the safety project changed
          sUdpVars.UnhandledReceivePacketCnt += 1;
        end_if;

      else
        // invalid command
        bd_LogRtMessagesInCy.UdpReceivedInvalidCommand := TRUE;
        sUdpVars.UnhandledReceivePacketCnt += 1;
      end_if;
    else
      // the only valid command here is the reinitialize or the confirmation for reinitialize
      if pPacketHeader^.Command = t_UdpCommand::UdpCmd_ReInitialize then
        // confirm the command and reinitialize
        sUdpVars.pTempSendBufferIRQ^.Header.Command            := t_UdpCommand::UdpCmd_ReInitConfirm;
        sUdpVars.pTempSendBufferIRQ^.Header.State              := t_UdpPacketHeaderV2.State.IsFromConsumer OR t_UdpPacketHeaderV2.State.IsFromProducer; // invalid state for normal data

        // only send command and state
        retcode := SendUDPData(sUdpVars.pTempSendBufferIRQ, sizeof(t_UdpPacketHeaderV2.Command) + sizeof(t_UdpPacketHeaderV2.State), udIPAddr);

        if retcode < 0 then
          sUdpVars.LastSendError := retcode;
          sUdpVars.SendErrorCnt += 1;
        else
          // remember the sender
          sUdpVars.ReInitSenderIP := udIPAddr;

          // reset module sync no (no more modules synchron)
          ModuleSyncNo := 0;

          // if sending the answer succeeded => reinitialize ourself
          ClassState := 0;

          // wait until we're synchron again
          InitSSW := _ClearRoutingInfos;

        end_if;

        b_AllLocalSlaveAddressesValid := FALSE;

      elsif pPacketHeader^.Command = t_UdpCommand::UdpCmd_ReInitConfirm then

        // we got this, finished with disconnecting this one
        if sUdpVars.ProducerConnectionNo then
          sUdpVars.paConnectionsToProducers^[sUdpVars.ProducerConnectionNo-1].WaitForResponse        := FALSE;
          sUdpVars.paConnectionsToProducers^[sUdpVars.ProducerConnectionNo-1].InfoBits.Disconnecting := FALSE;
        elsif sUdpVars.ConsumerConnectionNo then
          sUdpVars.paConnectionsToConsumers^[sUdpVars.ConsumerConnectionNo-1].WaitForResponse        := FALSE;
          sUdpVars.paConnectionsToConsumers^[sUdpVars.ConsumerConnectionNo-1].InfoBits.Disconnecting := FALSE;
          sUdpVars.paConnectionsToConsumers^[sUdpVars.ConsumerConnectionNo-1].bSequenceCntReceived   := FALSE; //reset flag to allow sequence counter for new udp communication
          sUdpVars.paConnectionsToConsumers^[sUdpVars.ConsumerConnectionNo-1].ActReceiveData.usHeaderVersion := 0;
          sUdpVars.paConnectionsToConsumers^[sUdpVars.ConsumerConnectionNo-1].ActSendData.usHeaderVersion    := 0;
        end_if;
      else
        // invalid state/command combination
        bd_LogRtMessagesInCy.UdpReceivedInvalidState := TRUE;
        sUdpVars.UnhandledReceivePacketCnt += 1;
      end_if;
    end_if;

  elsif pPacketHeader^.Command = t_UdpCommand::UdpCmd_ReInitialize then
    // before the clear config phase is finished, the only thing allowed is to answer on reinitialize requests (but without reinitializing again) or take the reinitconfirm packets

    // confirm the command and reinitialize
    sUdpVars.pTempSendBufferIRQ^.Header.Command            := t_UdpCommand::UdpCmd_ReInitConfirm;
    sUdpVars.pTempSendBufferIRQ^.Header.State              := t_UdpPacketHeaderV2.State.IsFromConsumer OR t_UdpPacketHeaderV2.State.IsFromProducer; // invalid state for normal data

    // only send command and state
    retcode := SendUDPData(sUdpVars.pTempSendBufferIRQ, sizeof(t_UdpPacketHeaderV2.Command) + sizeof(t_UdpPacketHeaderV2.State), udIPAddr);

    if retcode < 0 then
      sUdpVars.LastSendError := retcode;
      sUdpVars.SendErrorCnt += 1;
    end_if;

    b_AllLocalSlaveAddressesValid := FALSE;

  elsif pPacketHeader^.Command = t_UdpCommand::UdpCmd_ReInitConfirm then

    // we got this, finished with disconnecting this one
    if sUdpVars.ProducerConnectionNo then
      sUdpVars.paConnectionsToProducers^[sUdpVars.ProducerConnectionNo-1].WaitForResponse        := FALSE;
      sUdpVars.paConnectionsToProducers^[sUdpVars.ProducerConnectionNo-1].InfoBits.Disconnecting := FALSE;
      sUdpVars.paConnectionsToConsumers^[sUdpVars.ConsumerConnectionNo-1].ActReceiveData.usHeaderVersion := 0;
      sUdpVars.paConnectionsToConsumers^[sUdpVars.ConsumerConnectionNo-1].ActSendData.usHeaderVersion    := 0;
    elsif sUdpVars.ConsumerConnectionNo then
      sUdpVars.paConnectionsToConsumers^[sUdpVars.ConsumerConnectionNo-1].WaitForResponse        := FALSE;
      sUdpVars.paConnectionsToConsumers^[sUdpVars.ConsumerConnectionNo-1].InfoBits.Disconnecting := FALSE;
      sUdpVars.paConnectionsToConsumers^[sUdpVars.ConsumerConnectionNo-1].bSequenceCntReceived   := FALSE; //reset flag to allow sequence counter for new udp communication
      sUdpVars.paConnectionsToConsumers^[sUdpVars.ConsumerConnectionNo-1].ActReceiveData.usHeaderVersion := 0;
      sUdpVars.paConnectionsToConsumers^[sUdpVars.ConsumerConnectionNo-1].ActSendData.usHeaderVersion    := 0;
    end_if;

  end_if;

END_FUNCTION

FUNCTION SafetyManager::HandleUdpRequest
  VAR_INPUT
    pConnection 	: ^t_UdpConnection;
    pPacket 	: ^t_UdpPacketV1;
    udLength 	: UDINT;
  END_VAR
  VAR
    SequenceDifference : SINT;
  END_VAR

  if udLength >= (sizeof(pPacket^.Header)) then

    pConnection^.ReceivedPackages += 1;

    //Allow the sequence counter if it is a new udp communication.
    if pConnection^.bSequenceCntReceived = FALSE then
      //In order for the packet to be forwarded to safety, the sequencing counter must be reduced.
      pConnection^.ActReceiveData.usSequenceNumber:= pPacket^.Header.SequenceNumber-1;
      pConnection^.bSequenceCntReceived := TRUE;
    end_if;

    SequenceDifference$SINT := (pPacket^.Header.SequenceNumber$SINT - pConnection^.ActReceiveData.usSequenceNumber$SINT);

    // Only packages with a new or identical sequence counter are allowed.
    if (SequenceDifference >= 0) & (SequenceDifference < 127) then
      //set flag and timestamp for last request
      if pConnection^.WaitForResponse = TRUE then
        pConnection^.WaitForResponse := FALSE;
        pConnection^.LastResponseTime := ops.tAbsolute - pConnection^.TLastRequest;
        if pConnection^.LastResponseTime > pConnection^.MaxResponseTime then
          pConnection^.MaxResponseTime := pConnection^.LastResponseTime;
        end_if;
      end_if;

      //only forward data to safety if it is a new package
      if SequenceDifference > 0 then

        UdpReceiveData.SectionStart();
        // The data is only copied if more than 0 bytes are available in the package and the size is smaller then max size.
        if pPacket^.Header.PdoDataLength & pPacket^.Header.PdoDataLength <= UDP_MAX_PDO_SIZE then
          pConnection^.ActReceiveData.PdoLength := pPacket^.Header.PdoDataLength;
          _memcpy(ptr1:=#pConnection^.ActReceiveData.PdoData, ptr2:=#pPacket^.Data, cntr:=pConnection^.ActReceiveData.PdoLength);

          //check for communication ok of fsoe connection (CMD 0x64 = Connection)
          if pConnection^.ActReceiveData.PdoData[0] = 16#64 & pConnection^.bs_SingleLog.OldHeaderVersionOfResponseIF = FALSE then
            LogError("@04E1 (SafetyManager::HandleUdpRequest) [SL] The header version of the request interface doesn't support 4 byte sequence number!");
            LogValue("@04E1 (SafetyManager::HandleUdpRequest) [SL] IFCRC: 0x{0}, SafetyNbr: 0x{1}, IPAddress: 0x{2}", pConnection^.IFCRC, pConnection^.SafetyNbrOtherSide, pConnection^.IP);
            pConnection^.bs_SingleLog.OldHeaderVersionOfResponseIF := TRUE;
          end_if;
        else
          pConnection^.ActReceiveData.PdoLength := 0;
        end_if;

        if pPacket^.Header.SdoDataLength & (pConnection^.ActReceiveData.SdoLength = 0)
        & (pPacket^.Header.SdoDataLength <= UDP_MAX_SDO_SIZE) then
          pConnection^.ActReceiveData.SdoLength := pPacket^.Header.SdoDataLength;
          _memcpy(ptr1:=#pConnection^.ActReceiveData.SdoData, ptr2:=#pPacket^.Data + pConnection^.ActReceiveData.PdoLength, cntr:=pConnection^.ActReceiveData.SdoLength);
        end_if;
        UdpReceiveData.SectionStop();

      end_if;

      // save safety number of other side
      pConnection^.SafetyNbrOtherSide             := pPacket^.Header.SafetyNbr;
      pConnection^.ActReceiveData.usSequenceNumber:= pPacket^.Header.SequenceNumber;
      pConnection^.ActSendData.usSequenceNumber   := pConnection^.ActReceiveData.usSequenceNumber;
      //set sequence number of v2 header
      pConnection^.ActSendData.udSequenceNumber    := pConnection^.ActReceiveData.usSequenceNumber;
      pConnection^.ActReceiveData.udSequenceNumber := pConnection^.ActReceiveData.usSequenceNumber;

      //if the callback time is smaller than min request time and sequence diff = 0 its an old request -> don't send the response again
      if (ops.tAbsolute - pConnection^.TLastRequest) > UDP_MIN_REQUEST_TIME | SequenceDifference > 0 then
        pConnection^.SendResponse := TRUE;
      end_if;

    else
      //it's an old package
      sUdpVars.WrongSequenceInRequestCnt += 1;
      //if the last valid request is greater then maximal FSoE Watchdog Time we can reset the sequence Counter from this connection
      if (ops.tAbsolute - pConnection^.TLastRequest) > (UDP_DEFAULT_TRANSMISSION_TIME*2) then
        pConnection^.bSequenceCntReceived := FALSE;
//        pConnection^.TLastRequest := ops.tAbsolute;
      end_if;
    end_if;
  else
    sUdpVars.WrongReceiveUDPLength += 1;
  end_if;

END_FUNCTION

FUNCTION SafetyManager::HandleUdpRequestV2
  VAR_INPUT
    pConnection 	: ^t_UdpConnection;
    pPacket 	: ^t_UdpPacketV2;
    udLength 	: UDINT;
  END_VAR
  VAR
    SequenceDifference : DINT;
  END_VAR

  if udLength >= (sizeof(pPacket^.Header)) then

    pConnection^.ReceivedPackages += 1;

    //Allow the sequence counter if it is a new udp communication.
    if pConnection^.bSequenceCntReceived = FALSE then
      //In order for the packet to be forwarded to safety, the sequencing counter must be reduced.
      pConnection^.ActReceiveData.udSequenceNumber:= pPacket^.Header.SequenceNumber-1;
      pConnection^.bSequenceCntReceived := TRUE;
    end_if;

    SequenceDifference := pPacket^.Header.SequenceNumber$DINT - pConnection^.ActReceiveData.udSequenceNumber$DINT;

    // Only packages with a new or identical sequence counter are allowed.
    if (SequenceDifference >= 0) & (SequenceDifference < 127) then
      //set flag and timestamp for last request
      if pConnection^.WaitForResponse = TRUE then
        pConnection^.WaitForResponse := FALSE;
        pConnection^.LastResponseTime := ops.tAbsolute - pConnection^.TLastRequest;
        if pConnection^.LastResponseTime > pConnection^.MaxResponseTime then
          pConnection^.MaxResponseTime := pConnection^.LastResponseTime;
        end_if;
      end_if;

      //only forward data to safety if it is a new package
      if SequenceDifference > 0 then

        UdpReceiveData.SectionStart();
        // The data is only copied if more than 0 bytes are available in the package and the size is smaller then max size.
        if pPacket^.Header.PdoDataLength & pPacket^.Header.PdoDataLength <= UDP_MAX_PDO_SIZE then
          pConnection^.ActReceiveData.PdoLength := pPacket^.Header.PdoDataLength;
          _memcpy(ptr1:=#pConnection^.ActReceiveData.PdoData, ptr2:=#pPacket^.Data, cntr:=pConnection^.ActReceiveData.PdoLength);
        else
          pConnection^.ActReceiveData.PdoLength := 0;
        end_if;

        if pPacket^.Header.SdoDataLength & (pConnection^.ActReceiveData.SdoLength = 0)
        & (pPacket^.Header.SdoDataLength <= UDP_MAX_SDO_SIZE) then
          pConnection^.ActReceiveData.SdoLength := pPacket^.Header.SdoDataLength;
          _memcpy(ptr1:=#pConnection^.ActReceiveData.SdoData, ptr2:=#pPacket^.Data + pConnection^.ActReceiveData.PdoLength, cntr:=pConnection^.ActReceiveData.SdoLength);
        end_if;
        UdpReceiveData.SectionStop();

      end_if;

      // save safety number of other side
      pConnection^.SafetyNbrOtherSide             := pPacket^.Header.SafetyNbr;
      pConnection^.ActReceiveData.udSequenceNumber:= pPacket^.Header.SequenceNumber;
      pConnection^.ActSendData.udSequenceNumber   := pConnection^.ActReceiveData.udSequenceNumber;

      //if the callback time is smaller than min request time and sequence diff = 0 its an old request -> don't send the response again
      if (ops.tAbsolute - pConnection^.TLastRequest) > UDP_MIN_REQUEST_TIME | SequenceDifference > 0 then
        pConnection^.SendResponse := TRUE;
      end_if;

    else
      //it's an old package
      sUdpVars.WrongSequenceInRequestCnt += 1;
      //if the last valid request is greater then maximal FSoE Watchdog Time we can reset the sequence Counter from this connection
      if (ops.tAbsolute - pConnection^.TLastRequest) > (UDP_DEFAULT_TRANSMISSION_TIME*2) then
        pConnection^.bSequenceCntReceived := FALSE;
//        pConnection^.TLastRequest := ops.tAbsolute;
      end_if;
    end_if;
  else
    sUdpVars.WrongReceiveUDPLength += 1;
  end_if;

END_FUNCTION

FUNCTION SafetyManager::HandleUdpResponse
  VAR_INPUT
    pConnection 	: ^t_UdpConnection;
    pPacket 	: ^t_UdpPacketV1;
    udLength 	: UDINT;
  END_VAR
  VAR
    SequenceDifference : SINT;
  END_VAR

  //check length of udp data -> length must be more then header size
  if udLength >= (sizeof(pPacket^.Header)) then
    pConnection^.ReceivedPackages += 1;

    pConnection^.ActReceiveData.usSequenceNumber := pPacket^.Header.SequenceNumber;
    pConnection^.ActReceiveData.udSequenceNumber := pConnection^.ActReceiveData.usSequenceNumber;

    // Only packages with identical sequence counter are allowed.
    if pConnection^.ActReceiveData.usSequenceNumber = pConnection^.ActSendData.usSequenceNumber then
      // we got our response => increase the sequence number
      pConnection^.ActSendData.usSequenceNumber += 1;
      pConnection^.ActSendData.udSequenceNumber := pConnection^.ActSendData.usSequenceNumber;

      if pConnection^.WaitForResponse = TRUE then
        pConnection^.WaitForResponse := FALSE;
        pConnection^.LastResponseTime := ops.tAbsolute - pConnection^.TLastRequest;
        if pConnection^.LastResponseTime > pConnection^.MaxResponseTime then
          pConnection^.MaxResponseTime := pConnection^.LastResponseTime;
        end_if;
        pConnection^.TLastValidRequest := ops.tAbsolute;
      else
        sUdpVars.ReceivedUnexpectedResponse += 1;
        return;
      end_if;

      UdpReceiveData.SectionStart();

      // The data is only copied if more than 0 bytes are available in the package and the size is smaller then max size.
      if pPacket^.Header.PdoDataLength & pPacket^.Header.PdoDataLength <= UDP_MAX_PDO_SIZE then
        pConnection^.ActReceiveData.PdoLength := pPacket^.Header.PdoDataLength;
        _memcpy(ptr1:=#pConnection^.ActReceiveData.PdoData, ptr2:=#pPacket^.Data, cntr:=pConnection^.ActReceiveData.PdoLength);

        //check for communication ok of fsoe connection (CMD 0x64 = Connection)
        if pConnection^.ActReceiveData.PdoData[0] = 16#64 & pConnection^.bs_SingleLog.OldHeaderVersionOfResponseIF = FALSE then
          LogError("@04E0 (SafetyManager::HandleUdpResponse) The header version of the response interface doesn't support 4 byte sequence number!");
          LogValue("@04E1 (SafetyManager::HandleUdpResponse) [SL] IFCRC: 0x{0}, SafetyNbr: 0x{1}, IPAddress: 0x{2}", pConnection^.IFCRC, pConnection^.SafetyNbrOtherSide, pConnection^.IP);
          pConnection^.bs_SingleLog.OldHeaderVersionOfResponseIF := TRUE;
        end_if;
      else
        pConnection^.ActReceiveData.PdoLength := 0;
      end_if;

      if (pPacket^.Header.SdoDataLength) & (pConnection^.ActReceiveData.SdoLength = 0)
      & (pPacket^.Header.SdoDataLength <= UDP_MAX_SDO_SIZE) then
        pConnection^.ActReceiveData.SdoLength := pPacket^.Header.SdoDataLength;
        _memcpy(ptr1:=#pConnection^.ActReceiveData.SdoData, ptr2:=#pPacket^.Data + pConnection^.ActReceiveData.PdoLength, cntr:=pConnection^.ActReceiveData.SdoLength);
      end_if;

      UdpReceiveData.SectionStop();
    else
      //sequence counter is not the same
      sUdpVars.WrongSequenceInResponseCnt += 1;

      //check the sequence difference, it could be a retry from other side which contains sdo data
      SequenceDifference := pConnection^.ActReceiveData.udSequenceNumber$SINT - pConnection^.ActSendData.udSequenceNumber$SINT;

      UdpReceiveData.SectionStart();
      //if Sequence difference is -1 it could be a response retry with sdo data
      if (pPacket^.Header.SdoDataLength) & (pConnection^.ActReceiveData.SdoLength = 0)
      & (pPacket^.Header.SdoDataLength <= UDP_MAX_SDO_SIZE) & (SequenceDifference = -1) then
        pConnection^.ActReceiveData.SdoLength := pPacket^.Header.SdoDataLength;
        _memcpy(ptr1:=#pConnection^.ActReceiveData.SdoData, ptr2:=#pPacket^.Data + pConnection^.ActReceiveData.PdoLength, cntr:=pConnection^.ActReceiveData.SdoLength);
      end_if;
      UdpReceiveData.SectionStop();
    end_if;

    // save safety number of other side
    pConnection^.SafetyNbrOtherSide       := pPacket^.Header.SafetyNbr;
  else
    sUdpVars.WrongReceiveUDPLength += 1;
  end_if;

END_FUNCTION

FUNCTION SafetyManager::HandleUdpResponseV2
  VAR_INPUT
    pConnection 	: ^t_UdpConnection;
    pPacket 	: ^t_UdpPacketV2;
    udLength 	: UDINT;
  END_VAR
  VAR
    SequenceDifference : DINT;
  END_VAR

  //check length of udp data -> length must be more then header size
  if udLength >= (sizeof(pPacket^.Header)) then

    pConnection^.ReceivedPackages += 1;
    pConnection^.ActReceiveData.udSequenceNumber := pPacket^.Header.SequenceNumber;

    // Only packages with identical sequence counter are allowed.
    if pConnection^.ActReceiveData.udSequenceNumber = pConnection^.ActSendData.udSequenceNumber then
      // we got our response => increase the sequence number
      pConnection^.ActSendData.udSequenceNumber += 1;

      if pConnection^.WaitForResponse = TRUE then
        pConnection^.WaitForResponse := FALSE;
        pConnection^.LastResponseTime := ops.tAbsolute - pConnection^.TLastRequest;
        if pConnection^.LastResponseTime > pConnection^.MaxResponseTime then
          pConnection^.MaxResponseTime := pConnection^.LastResponseTime;
        end_if;
        pConnection^.TLastValidRequest := ops.tAbsolute;
      else
        sUdpVars.ReceivedUnexpectedResponse += 1;
        return;
      end_if;

      UdpReceiveData.SectionStart();

      // The data is only copied if more than 0 bytes are available in the package and the size is smaller then max size.
      if pPacket^.Header.PdoDataLength & pPacket^.Header.PdoDataLength <= UDP_MAX_PDO_SIZE then
        pConnection^.ActReceiveData.PdoLength := pPacket^.Header.PdoDataLength;
        _memcpy(ptr1:=#pConnection^.ActReceiveData.PdoData, ptr2:=#pPacket^.Data, cntr:=pConnection^.ActReceiveData.PdoLength);
      else
        pConnection^.ActReceiveData.PdoLength := 0;
      end_if;

      if (pPacket^.Header.SdoDataLength) & (pConnection^.ActReceiveData.SdoLength = 0)
      & (pPacket^.Header.SdoDataLength <= UDP_MAX_SDO_SIZE) then
        pConnection^.ActReceiveData.SdoLength := pPacket^.Header.SdoDataLength;
        _memcpy(ptr1:=#pConnection^.ActReceiveData.SdoData, ptr2:=#pPacket^.Data + pConnection^.ActReceiveData.PdoLength, cntr:=pConnection^.ActReceiveData.SdoLength);
      end_if;

      UdpReceiveData.SectionStop();
    else
      //sequence counter is not the same
      sUdpVars.WrongSequenceInResponseCnt += 1;

      //check the sequence difference, it could be a retry from other side which contains sdo data
      SequenceDifference := pConnection^.ActReceiveData.udSequenceNumber$DINT - pConnection^.ActSendData.udSequenceNumber$DINT;

      UdpReceiveData.SectionStart();
      //if Sequence difference is -1 it could be a response retry with sdo data
      if (pPacket^.Header.SdoDataLength) & (pConnection^.ActReceiveData.SdoLength = 0)
      & (pPacket^.Header.SdoDataLength <= UDP_MAX_SDO_SIZE) & (SequenceDifference = -1) then
        pConnection^.ActReceiveData.SdoLength := pPacket^.Header.SdoDataLength;
        _memcpy(ptr1:=#pConnection^.ActReceiveData.SdoData, ptr2:=#pPacket^.Data + pConnection^.ActReceiveData.PdoLength, cntr:=pConnection^.ActReceiveData.SdoLength);
      end_if;
      UdpReceiveData.SectionStop();
    end_if;

    // save safety number of other side
    pConnection^.SafetyNbrOtherSide       := pPacket^.Header.SafetyNbr;
  else
    sUdpVars.WrongReceiveUDPLength += 1;
  end_if;

END_FUNCTION

FUNCTION SafetyManager::ForwardReceivedUdpSDOs
  VAR_INPUT
    paConnections 	: ^t_aUdpConnections;
    ConnectionNo 	: UDINT;
  END_VAR
  VAR
    i               : UDINT;
    pActConnection  : ^t_UdpConnection;
    pHelpCfg        : ^t_CfgListElem;
    pHelpModule     : ^t_ModuleListElem;
    InterfaceCRC    : HDINT;
    SafetyNumber    : HDINT;
    MyPara          : CmdStruct;
    MyResult        : results;
    pDO 	          : ^SafetyCDIAS_Base::SDOHeader;
    pCompDestPath   : ^USINT;
    pHelpSafety     : ^t_SafetyComponent;
    ResponseValue   : BOOL;
    FoundTarget     : BOOL;
  END_VAR

  ResponseValue := paConnections = sUdpVars.paConnectionsToProducers;

  pActConnection := #paConnections^[0];
  for i := 0 to (ConnectionNo-1) do

    // check if there is a SDO to forward
    if pActConnection^.ActReceiveData.SdoLength then

      FoundTarget := FALSE;

      UdpReceiveData.SectionStart();

      // get a pointer to the compressed destination path
      pDO := (#pActConnection^.ActReceiveData.SdoData)$^SafetyCDIAS_Base::SDOHeader;
      if (pDO^.StdHeader.Typ.Response = ResponseValue) then
        pCompDestPath := (#pDO^.DstAdr)$^USINT;

        // check if it's addressed by topology path and it's an IP
        if ((pDO^.StdHeader.Typ AND SSDO_MASK_TYPE) = FRM_TYPECODE_SSDO_MOD_TP) & (pCompDestPath^ = INTERFACE_IP_MODE) then
          // after the mode byte we find the interface CRC
          InterfaceCRC := ((pCompDestPath + 1)$^HDINT)^;

          // search all configs, all moduleconfigs

          pHelpCfg := pConfigs;
          while pHelpCfg & pActConnection^.ActReceiveData.SdoLength do
            pHelpModule := pHelpCfg^.pFirstModuleCfg;
            while pHelpModule & pActConnection^.ActReceiveData.SdoLength do
              if pHelpModule^.ModuleInfo.InterfaceCRC = InterfaceCRC then
                // we found the interface CRC, now we have to make a connection via the SafetyNumber between the actual module config and the module handles
                pHelpSafety := pFirstSafetyComponent;
                while pHelpSafety & pActConnection^.ActReceiveData.SdoLength do
                  // we compare the safety number
                  if pHelpSafety^.SafetyNbr = pHelpModule^.ModuleInfo.SafetyNbr then

                    MyPara.uiCmd := CMD_SM_SDO_TO_MODULE;
                    MyPara.aPara[0] := pActConnection^.ActReceiveData.SdoLength;
                    MyPara.aPara[1] := (#pActConnection^.ActReceiveData.SdoData)$DINT;
                    MyPara.aPara[2] := this$DINT;

                    pHelpSafety^.pThis^.NewInst(#MyPara, #MyResult);

                    FoundTarget := TRUE;
                  end_if;

                  pHelpSafety := pHelpSafety^.pNext;
                end_while;
              end_if;

              pHelpModule := pHelpModule^.pNext;
            end_while;

            pHelpCfg := pHelpCfg^.pNext;
          end_while;
        else
          SafetyNumber := pDO^.DstAdr;

          // search by safety number and forward to internal module
          pHelpSafety := pFirstSafetyComponent;
          while pHelpSafety & pActConnection^.ActReceiveData.SdoLength do
            // we compare the safety number
            if pHelpSafety^.SafetyNbr = SafetyNumber then
              MyPara.uiCmd := CMD_SM_SDO_TO_MODULE;
              MyPara.aPara[0] := pActConnection^.ActReceiveData.SdoLength;
              MyPara.aPara[1] := (#pActConnection^.ActReceiveData.SdoData)$DINT;
              MyPara.aPara[2] := this$DINT;

              pHelpSafety^.pThis^.NewInst(#MyPara, #MyResult);

              FoundTarget := TRUE;
            end_if;

            pHelpSafety := pHelpSafety^.pNext;
          end_while;
        end_if;

        // reset length if the response bit matches (if we found it, we already forwarded it. if not, we're not going to find it next time)
        pActConnection^.ActReceiveData.SdoLength := 0;
      else
        // check which list it is
        if ResponseValue then
          sUdpVars.InvalidResponseSettingAtFowardingProducerList += 1;
        else
          sUdpVars.InvalidResponseSettingAtFowardingConsumerList += 1;
        end_if;
      end_if;

      UdpReceiveData.SectionStop();

    end_if;

    pActConnection += sizeof(t_UdpConnection);
  end_for;

END_FUNCTION

FUNCTION SafetyManager::ForwardSDO2UdpBySafetyNbr
  VAR_INPUT
    SDOLength 	: UINT;
    pSDO 	: ^USINT;
  END_VAR
  VAR_OUTPUT
    FoundTarged 	: BOOL;
  END_VAR
  VAR
    i               : UDINT;
    pActConnection  : ^t_UdpConnection;
    TargetSafetyNbr : HDINT;
    pDO 	          : ^SafetyCDIAS_Base::SDOHeader;
  END_VAR

  FoundTarged := FALSE;

  // get a pointer to the compressed destination path
  pDO := pSDO$^SafetyCDIAS_Base::SDOHeader;
  TargetSafetyNbr := pDO^.DstAdr;

  if sUdpVars.ConsumerConnectionNo then
    pActConnection := #sUdpVars.paConnectionsToConsumers^[0];
    for i := 0 to (sUdpVars.ConsumerConnectionNo-1) do
      // the safety number has to match and since it's a message to a consumer it has to be a response
      if (pActConnection^.SafetyNbrOtherSide = TargetSafetyNbr) & (pDO^.StdHeader.Typ.Response = TRUE) then
        // got it => forward the SDO
        if SDOLength <= UDP_MAX_SDO_SIZE then
          // check for unsent SDO first
          if pActConnection^.ActSendData.SdoLength = 0 then
            UdpSendData.SectionStart();

            _memcpy(ptr1:=#pActConnection^.ActSendData.SdoData, ptr2:=pSDO, cntr:=SDOLength);
            pActConnection^.ActSendData.SdoLength     := SDOLength$USINT;

            UdpSendData.SectionStop();
          else
            sUdpVars.SdoAlreadyUsedCnt += 1;
          end_if;
        else
          LogError("@046E (SafetyManager::ForwardSDO2UdpBySafetyNbr) SDO size exceeds the allowed size (Compressed Topology Path: UDP)");
        end_if;

        FoundTarged := TRUE;
        return;
      end_if;

      pActConnection += sizeof(t_UdpConnection);
    end_for;
  end_if;

  if sUdpVars.ProducerConnectionNo then
    pActConnection := #sUdpVars.paConnectionsToProducers^[0];
    for i := 0 to (sUdpVars.ProducerConnectionNo-1) do
      // the safety number has to match and since it's a message to a producer it has to be a request
      if (pActConnection^.SafetyNbrOtherSide = TargetSafetyNbr) & (pDO^.StdHeader.Typ.Response = FALSE) then
        // got it => forward the SDO
        if SDOLength <= UDP_MAX_SDO_SIZE then
          // check for unsent SDO first
          if pActConnection^.ActSendData.SdoLength = 0 then
            UdpSendData.SectionStart();

            _memcpy(ptr1:=#pActConnection^.ActSendData.SdoData, ptr2:=pSDO, cntr:=SDOLength);
            pActConnection^.ActSendData.SdoLength     := SDOLength$USINT;

            UdpSendData.SectionStop();
          else
            sUdpVars.SdoAlreadyUsedCnt += 1;
          end_if;
        else
          LogError("@046E (SafetyManager::ForwardSDO2Udp) SDO size exceeds the allowed size (Compressed Topology Path: UDP)");
        end_if;

        FoundTarged := TRUE;
        return;
      end_if;

      pActConnection += sizeof(t_UdpConnection);
    end_for;
  end_if;

END_FUNCTION

FUNCTION SafetyManager::ShareUdpConnectionInfos
  VAR
    i                 : UDINT;
    pUdpConnection    : ^t_UdpConnection;
    AnythingMissing   : BOOL;
    ActInitialized    : BOOL;
    FoundConnection   : BOOL;
    pHelpSafety       : ^t_SafetyComponent;
    pHelpCfg          : ^t_CfgListElem;
    pFSoEConnection   : ^t_FSoEConnectionDetails;
    MyPara            : CmdStruct;
    MyResult          : results;
    retcode           : iprStates;

    ModuleReadOffset  : UINT;
    ModuleReadSize    : UINT;
    ModuleWriteOffset : UINT;
    ModuleWriteSize   : UINT;
    MngReadOffset     : UINT;
    MngReadSize       : UINT;
    MngWriteOffset    : UINT;
    MngWriteSize      : UINT;
  END_VAR

  AnythingMissing := FALSE;

  if sUdpVars.ConsumerConnectionNo then
    pUdpConnection := #sUdpVars.paConnectionsToConsumers^[0];
    for i := 0 to (sUdpVars.ConsumerConnectionNo-1) do
      // check if we received something so far at this connection
      if (pUdpConnection^.ReceivedPackages & (pUdpConnection^.InfoBits.PdosInitialized = FALSE)) then
        FoundConnection := ActInitialized := FALSE;

        // check FSoE Connections in the available configs if there is a match at the interface CRC
        pHelpCfg := pConfigs;
        while pHelpCfg & (FoundConnection = FALSE) do
          pFSoEConnection := pHelpCfg^.pFirstFSoEConnection;
          while pFSoEConnection & (FoundConnection = FALSE) do
            // only interface slave connections which are not used yet are relevant
            if pFSoEConnection^.Flags.IsInterfaceConnection & (pFSoEConnection^.Flags.IsMaster = FALSE) & (pFSoEConnection^.InternalConnectionState = FCS_RESET) &
               pFSoEConnection^.pSlavePathComp & ((pFSoEConnection^.pSlavePathComp$^HDINT + 1)^ = pUdpConnection^.IFCRC) then

              // found the connection
              FoundConnection := TRUE;

              // now try to initialize it

              pHelpSafety := pFirstSafetyComponent;
              while pHelpSafety do
                if pHelpSafety^.SafetyNbr = pFSoEConnection^.OwnerSafetyNbr then
                  exit;
                end_if;

                pHelpSafety := pHelpSafety^.pNext;
              end_while;

              if pHelpSafety then
#ifdef SAFETY_DEBUG_LOGGING_ACTIVATED
#pragma message("RamAnd 20.11.2014 16:41 \ testweise mapping loggen")
                LogValue("@DBG (SafetyManager::ShareUdpConnectionInfos) <This side is Slave> ConnectionID: 0x{0}, SlaveAddress: 0x{1}, IFCRC: 0x{2}", Value:=pFSoEConnection^.ConnectionID, Value2:=pFSoEConnection^.SlaveAddress, Value3 := (pFSoEConnection^.pSlavePathComp$^HDINT + 1)^);
                LogValue("@DBG (SafetyManager::ShareUdpConnectionInfos) <This side is Slave> UdpInfo: SNr: 0x{0}, SNrOtherSide: 0x{1}, IFCRC: 0x{2}", Value:=pUdpConnection^.SafetyNbr, Value2:=pUdpConnection^.SafetyNbrOtherSide, Value3 := pUdpConnection^.IFCRC);
#endif

                // the module is slave and the managing module master
                ModuleReadOffset  := pFSoEConnection^.SlaveReadOffset;
                ModuleReadSize    := pFSoEConnection^.MasterWriteSize;
                ModuleWriteOffset := pFSoEConnection^.SlaveWriteOffset;
                ModuleWriteSize   := pFSoEConnection^.MasterReadSize;
                MngReadOffset     := 0; // offsets in managing modules are always dynamic
                MngReadSize       := pFSoEConnection^.MasterReadSize;
                MngWriteOffset    := 0; // offsets in managing modules are always dynamic
                MngWriteSize      := pFSoEConnection^.MasterWriteSize;

#ifdef SAFETY_DEBUG_LOGGING_ACTIVATED
#pragma message("RamAnd 20.11.2014 16:41 \ testweise mapping loggen")
                LogValue("@DBG (SafetyManager::ShareUdpConnectionInfos) Modul => Udp: Rd Offset Modul: 0x{0}, IP: 0x{1}, Größe: 0x{2}", Value:=ModuleReadOffset, Value2:=pUdpConnection^.IP, Value3:=ModuleReadSize);
#endif

                MyPara.uiCmd    := CMD_SM_ADD_INPUT_PDO;
                MyPara.aPara[0] := (#pUdpConnection^.ThreadSafePdoReceiveBuffer)$DINT;
                MyPara.aPara[1] := 0;
                MyPara.aPara[2] := pUdpConnection^.SafetyNbrOtherSide$DINT;
                MyPara.aPara[3] := ModuleWriteSize;
                MyPara.aPara[4] := 0;
                MyPara.aPara[5] := 0;
                MyPara.aPara[6] := 0;
                MyPara.aPara[7] := ModuleWriteOffset;
                MyPara.aPara[8] := SM_IF_VALIDITY_MARK$DINT;
                MyPara.aPara[9] := TRUE;

                retcode := pHelpSafety^.pThis^.NewInst(#MyPara, #MyResult);

                if retcode = ERROR then
                  LogError("@0848 (SafetyManager::ShareUdpConnectionInfos) Failed to add input PDO for a connection to a Consumer");

                  // mark the connection to not try again later
                  pFSoEConnection^.InternalConnectionState := FCS_NOT_INITIALIZED;

                  return;
                elsif retcode = BUSY then
                  // try again later (skip further initialisation steps)
                  return;
                end_if;

                if FSoEInputPDONo < MAX_FSOE_CONNECTIONS then
                  aFSoEInputPDOs[FSoEInputPDONo].pSafety    := pHelpSafety;
                  aFSoEInputPDOs[FSoEInputPDONo].pMem       := MyPara.aPara[0];
                  FSoEInputPDONo                            += 1;

                  pUdpConnection^.ActReceiveData.PdoLength  := ModuleWriteSize;
                else
                  LogValue("@0490 (SafetyManager::ShareUdpConnectionInfos) Maximum limit of allowed FSoE input Frames exceeded (0x{0})", Value:=MAX_FSOE_CONNECTIONS);
                  exit;
                end_if;

                if sUdpVars.ReceiveCopyCmdNo < MAX_UDP_IF_ALLOWED then
                  sUdpVars.aReceiveCopyCmds[sUdpVars.ReceiveCopyCmdNo].pSource      := (#pUdpConnection^.ActReceiveData.PdoData)$^USINT;
                  sUdpVars.aReceiveCopyCmds[sUdpVars.ReceiveCopyCmdNo].pDest        := MyPara.aPara[0]$^USINT;
                  sUdpVars.aReceiveCopyCmds[sUdpVars.ReceiveCopyCmdNo].Size         := ModuleWriteSize;
                  sUdpVars.ReceiveCopyCmdNo                                            += 1;
                else
                  LogValue("@049F (SafetyManager::ShareUdpConnectionInfos) Maximum limit of allowed UDP receive copy commands exceeded (0x{0})", Value:=MAX_UDP_IF_ALLOWED);
                  exit;
                end_if;

                MyPara.uiCmd    := CMD_SM_ADD_OUTPUT_PDO;
                MyPara.aPara[0] := 1;  // mark as interface frame PDO
                pHelpSafety^.pThis^.NewInst(#MyPara, #MyResult);

//                  pPDOElement^.SourceInfo.pPDOMem       := MyResult.aData[0]$^USINT;
//                  pPDOElement^.SourceInfo.pPDOMemDPRAM  := MyResult.aData[4]$^USINT;
//                  pPDOElement^.SourceInfo.HandlePDODPRAM:= MyResult.aData[8]$UDINT;   // Needed for Payload Support
//                  pPDOElement^.SourceInfo.OffsetPDODPRAM:= MyResult.aData[12]$UDINT;  // Needed for Payload Support

                if sUdpVars.SendCopyCmdNo < MAX_UDP_IF_ALLOWED then
                  sUdpVars.aSendCopyCmds[sUdpVars.SendCopyCmdNo].pSource      := MyResult.aData[0]$^USINT + ModuleReadOffset;
                  sUdpVars.aSendCopyCmds[sUdpVars.SendCopyCmdNo].pDest        := #pUdpConnection^.ActSendData.PdoData;
                  sUdpVars.aSendCopyCmds[sUdpVars.SendCopyCmdNo].Size         := ModuleReadSize;
                  sUdpVars.SendCopyCmdNo                                         += 1;

                  pUdpConnection^.ActSendData.PdoLength           := ModuleReadSize;
                else
                  LogValue("@049E (SafetyManager::ShareUdpConnectionInfos) Maximum limit of allowed UDP send copy commands exceeded (0x{0})", Value:=MAX_UDP_IF_ALLOWED);
                  exit;
                end_if;

#ifdef SAFETY_DEBUG_LOGGING_ACTIVATED
#pragma message("RamAnd 20.11.2014 16:41 \ testweise mapping loggen")
                LogValue("@DBG (SafetyManager::ShareUdpConnectionInfos) Udp => Modul: Wr Offset Modul: 0x{0}, IP: 0x{1}, Größe: 0x{2}", Value:=ModuleWriteOffset, Value2:=pUdpConnection^.IP, Value3:=ModuleWriteSize);
#endif

                // mark the FSoE connection as established
                pFSoEConnection^.InternalConnectionState  := FCS_CONNECTION;

                // mark the udp connection as established
                pUdpConnection^.InfoBits.PdosInitialized  := TRUE;

                // connection initialized
                ActInitialized                            := TRUE;

                // check if we have all slave addresses now
                CheckLocalSlaveAddresses();
              else
                LogValue("@495 (SafetyManager::ShareUdpConnectionInfos) Could not find safety module with safety number 0x{0} for FSoE interface connection", Value:=pFSoEConnection^.OwnerSafetyNbr);
              end_if;
            end_if;

            pFSoEConnection := pFSoEConnection^.pNext;
          end_while;

          if pHelpCfg then
            pHelpCfg := pHelpCfg^.pNext;
          end_if;
        end_while;

        if ActInitialized = FALSE then
          AnythingMissing := TRUE;
        end_if;
      elsif (pUdpConnection^.ReceivedPackages = 0) then
        AnythingMissing := TRUE;
      end_if;

      pUdpConnection += sizeof(t_UdpConnection);
    end_for;
  end_if;

  if sUdpVars.ProducerConnectionNo then
    pUdpConnection := #sUdpVars.paConnectionsToProducers^[0];
    for i := 0 to (sUdpVars.ProducerConnectionNo-1) do
      // check if we received something so far at this connection
      if (pUdpConnection^.ReceivedPackages & (pUdpConnection^.InfoBits.PdosInitialized = FALSE)) then
        FoundConnection := ActInitialized := FALSE;

        // check FSoE Connections in the available configs if there is a match at the interface CRC
        pHelpCfg := pConfigs;
        while pHelpCfg & (FoundConnection = FALSE) do
          pFSoEConnection := pHelpCfg^.pFirstFSoEConnection;
          while pFSoEConnection & (FoundConnection = FALSE) do
            // only interface master connections which are not used are relevant
            if pFSoEConnection^.Flags.IsInterfaceConnection & pFSoEConnection^.Flags.IsMaster & (pFSoEConnection^.InternalConnectionState = FCS_RESET) then
              // check if it's our connection
              if ( pFSoEConnection^.pSlavePathComp) &
                 ( pFSoEConnection^.pSlavePathComp^             = INTERFACE_IP_MODE) &
                 ((pFSoEConnection^.pSlavePathComp$^HDINT + 1)^ = pUdpConnection^.IFCRC) &
                 ((pFSoEConnection^.pSlavePathComp$^HDINT + 5)^ = pUdpConnection^.IP) then

                // found the connection
                FoundConnection := TRUE;

                // now try to initialize it

                pHelpSafety := pFirstSafetyComponent;
                while pHelpSafety do
                  if pHelpSafety^.SafetyNbr = pFSoEConnection^.OwnerSafetyNbr then
                    exit;
                  end_if;

                  pHelpSafety := pHelpSafety^.pNext;
                end_while;

                if pHelpSafety then
  #ifdef SAFETY_DEBUG_LOGGING_ACTIVATED
  #pragma message("RamAnd 20.11.2014 16:41 \ testweise mapping loggen")
                  LogValue("@DBG (SafetyManager::ShareUdpConnectionInfos) <This side is Master> ConnectionID: 0x{0}, SlaveAddress: 0x{1}, InterfaceCRC: 0x{2}", Value:=pFSoEConnection^.ConnectionID, Value2:=pFSoEConnection^.SlaveAddress, Value3 := pUdpConnection^.IFCRC);
#endif

                  // the module is master and the managing module slave
                  ModuleReadOffset  := pFSoEConnection^.MasterReadOffset;
                  ModuleReadSize    := pFSoEConnection^.MasterReadSize;
                  ModuleWriteOffset := pFSoEConnection^.MasterWriteOffset;
                  ModuleWriteSize   := pFSoEConnection^.MasterWriteSize;
                  MngReadOffset     := 0; // offsets in managing modules are always dynamic
                  MngReadSize       := pFSoEConnection^.MasterWriteSize;
                  MngWriteOffset    := 0; // offsets in managing modules are always dynamic
                  MngWriteSize      := pFSoEConnection^.MasterReadSize;

  #ifdef SAFETY_DEBUG_LOGGING_ACTIVATED
  #pragma message("RamAnd 20.11.2014 16:41 \ testweise mapping loggen")
                  LogValue("@DBG (SafetyManager::ShareUdpConnectionInfos) Modul => Udp: Rd Offset Modul: 0x{0}, IP: 0x{1}, Größe: 0x{2}", Value:=ModuleReadOffset, Value2:=pUdpConnection^.IP, Value3:=ModuleReadSize);
  #endif

                  MyPara.uiCmd    := CMD_SM_ADD_INPUT_PDO;
                  MyPara.aPara[0] := (#pUdpConnection^.ThreadSafePdoReceiveBuffer)$DINT;
                  MyPara.aPara[1] := 0;
                  MyPara.aPara[2] := pUdpConnection^.SafetyNbrOtherSide$DINT;
                  MyPara.aPara[3] := ModuleWriteSize;
                  MyPara.aPara[4] := 0;
                  MyPara.aPara[5] := 0;
                  MyPara.aPara[6] := 0;
                  MyPara.aPara[7] := ModuleWriteOffset;
                  MyPara.aPara[8] := SM_IF_VALIDITY_MARK$DINT;
                  MyPara.aPara[9] := TRUE;

                  retcode := pHelpSafety^.pThis^.NewInst(#MyPara, #MyResult);

                  if retcode = ERROR then
                    LogError("@0849 (SafetyManager::ShareUdpConnectionInfos) Failed to add input PDO for a connection to a Producer");

                    // mark the connection to not try again later
                    pFSoEConnection^.InternalConnectionState := FCS_NOT_INITIALIZED;

                    return;
                  elsif retcode = BUSY then
                    // try again later (skip further initialisation steps)
                    return;
                  end_if;

                  if FSoEInputPDONo < MAX_FSOE_CONNECTIONS then
                    aFSoEInputPDOs[FSoEInputPDONo].pSafety    := pHelpSafety;
                    aFSoEInputPDOs[FSoEInputPDONo].pMem       := MyPara.aPara[0];
                    FSoEInputPDONo += 1;

                    pUdpConnection^.ActReceiveData.PdoLength  := ModuleWriteSize;
                  else
                    LogValue("@0490 (SafetyManager::ShareUdpConnectionInfos) Maximum limit of allowed FSoE input Frames exceeded (0x{0})", Value:=MAX_FSOE_CONNECTIONS);
                    exit;
                  end_if;

                  if sUdpVars.ReceiveCopyCmdNo < MAX_UDP_IF_ALLOWED then
                    sUdpVars.aReceiveCopyCmds[sUdpVars.ReceiveCopyCmdNo].pSource  := (#pUdpConnection^.ActReceiveData.PdoData)$^USINT;
                    sUdpVars.aReceiveCopyCmds[sUdpVars.ReceiveCopyCmdNo].pDest    := MyPara.aPara[0]$^USINT;
                    sUdpVars.aReceiveCopyCmds[sUdpVars.ReceiveCopyCmdNo].Size     := ModuleWriteSize;
                    sUdpVars.ReceiveCopyCmdNo                                        += 1;
                  else
                    LogValue("@049F (SafetyManager::ShareUdpConnectionInfos) Maximum limit of allowed UDP receive copy commands exceeded (0x{0})", Value:=MAX_UDP_IF_ALLOWED);
                    exit;
                  end_if;

                  MyPara.uiCmd      := CMD_SM_ADD_OUTPUT_PDO;
                  MyPara.aPara[0]   := 1;  // mark as interface frame PDO
                  pHelpSafety^.pThis^.NewInst(#MyPara, #MyResult);

  //                  pPDOElement^.SourceInfo.pPDOMem       := MyResult.aData[0]$^USINT;
  //                  pPDOElement^.SourceInfo.pPDOMemDPRAM  := MyResult.aData[4]$^USINT;
  //                  pPDOElement^.SourceInfo.HandlePDODPRAM:= MyResult.aData[8]$UDINT;   // Needed for Payload Support
  //                  pPDOElement^.SourceInfo.OffsetPDODPRAM:= MyResult.aData[12]$UDINT;  // Needed for Payload Support

                  if sUdpVars.SendCopyCmdNo < MAX_UDP_IF_ALLOWED then
                    sUdpVars.aSendCopyCmds[sUdpVars.SendCopyCmdNo].pSource      := MyResult.aData[0]$^USINT + ModuleReadOffset;
                    sUdpVars.aSendCopyCmds[sUdpVars.SendCopyCmdNo].pDest        := #pUdpConnection^.ActSendData.PdoData;
                    sUdpVars.aSendCopyCmds[sUdpVars.SendCopyCmdNo].Size         := ModuleReadSize;
                    sUdpVars.SendCopyCmdNo                                         += 1;

                    pUdpConnection^.ActSendData.PdoLength                             := ModuleReadSize;
                  else
                    LogValue("@049E (SafetyManager::ShareUdpConnectionInfos) Maximum limit of allowed UDP send copy commands exceeded (0x{0})", Value:=MAX_UDP_IF_ALLOWED);
                    exit;
                  end_if;

  #ifdef SAFETY_DEBUG_LOGGING_ACTIVATED
  #pragma message("RamAnd 20.11.2014 16:41 \ testweise mapping loggen")
                  LogValue("@DBG (SafetyManager::ShareUdpConnectionInfos) Udp => Modul: Wr Offset Modul: 0x{0}, IP: 0x{1}, Größe: 0x{2}", Value:=ModuleWriteOffset, Value2:=pUdpConnection^.IP, Value3:=ModuleWriteSize);
  #endif

                  // mark the FSoE connection as established
                  pFSoEConnection^.InternalConnectionState  := FCS_CONNECTION;

                  // mark the udp connection as established
                  pUdpConnection^.InfoBits.PdosInitialized  := TRUE;

                  // connection initialized
                  ActInitialized                            := TRUE;

                  // check if we have all slave addresses now
                  CheckLocalSlaveAddresses();
                else
                  LogValue("@0495 (SafetyManager::ShareUdpConnectionInfos) Could not find safety module with safety number 0x{0} for FSoE interface connection", Value:=pFSoEConnection^.OwnerSafetyNbr);
                end_if;

              end_if;

            end_if;

            pFSoEConnection := pFSoEConnection^.pNext;
          end_while;

          pHelpCfg := pHelpCfg^.pNext;
       end_while;

        if ActInitialized = FALSE then
          AnythingMissing := TRUE;
        end_if;
      elsif (pUdpConnection^.ReceivedPackages = 0) then
        AnythingMissing := TRUE;
      end_if;

      pUdpConnection += sizeof(t_UdpConnection);
    end_for;
  end_if;

  // if all available udp connections are initialized => set the marker for not coming here any more
  if AnythingMissing = FALSE then
    sUdpVars.ConnectionsInitialized := TRUE;

    // update scheduler grid
    SetUdpSchedulerGrid();
  end_if;

END_FUNCTION

FUNCTION SafetyManager::SetUdpSchedulerGrid
  VAR
    Temp            : UDINT;
    bGetRequestTimeout : BOOL;
  END_VAR

  bGetRequestTimeout := FALSE;

  // we can only calculate if there are producer connections => otherwise the scheduler is not active
  if sUdpVars.ProducerConnectionNo then

    // the timeout is calculated so we could fit 4 timed out transmissions into the watchdog time (watchdog = 2*transmission time)
    Temp := sUdpVars.LowestTransmissionTime_ms * 2 / 4;

    // if the result is smaller than the minimum timeout => set it to the minimum
    if Temp < UDP_MIN_REQUEST_TIMEOUT then
      Temp := UDP_MIN_REQUEST_TIMEOUT;
    end_if;
